(* IEC 61131-3 sources: plc-st-coding-agent/progress/evidence/f14_v10_full_20261113/jobs/codex_minimax-m27 (part 7) *)

(* ---- self-hard-06.candidate_02.st ---- *)
The error is on line 65: assigning WORD to BOOL. Let me fix the `tmpTwoAgoPrevCond` variable and the consecutive 3-scan tracking logic.
FUNCTION_BLOCK FB
VAR_INPUT
    runRequest      : BOOL;
    pressure        : REAL;
    pressureValid   : BOOL;
    fuelFlow        : REAL;
    steamFlow       : REAL;
    outletCmd       : INT;
    outletFeedback  : INT;
    resetBtn        : BOOL;
END_VAR
VAR_OUTPUT
    tripLatched     : BOOL;
    fuelPermit      : BOOL;
    currentCauseMask: WORD;
    latchedCauseMask: WORD;
    diagnosticActive: BOOL;
END_VAR
VAR
    prevResetBtn            : BOOL := FALSE;
    prevRunRequest          : BOOL := FALSE;
    prevPressureValid       : BOOL := FALSE;
    prevPressure            : REAL := 0.0;
    prevOutletCmd           : INT := 0;
    prevOutletFeedback      : INT := 0;
    prevTripLatched         : BOOL := FALSE;
    prevCurrentCauseMask    : WORD := 0;
    prevLatchedCauseMask    : WORD := 0;
    prevStuckCond           : BOOL := FALSE;
    prev2StuckCond          : BOOL := FALSE;
    tmpRisingReset          : BOOL;
    tmpStuckCond            : BOOL;
    tmpCurrentMask          : WORD;
    tmpOverpressureValid    : BOOL;
END_VAR

(* CONTRACT:
   | Output/State    | Activation         | Retention       | Reset/Deactivation           | Same-scan Priority | Units/Boundaries       |
   |-----------------|--------------------|-----------------|-------------------------------|--------------------|------------------------|
   | tripLatched     | runRequest & (!pressureValid OR pressure>=4500.0) | Hold until resetBtn rising & !runRequest & pressureValid & pressure<=4200.0 | resetBtn rising edge clears | Same-scan with clue calc | BOOL; 4500/4200 kPa hysteresis |
   | fuelPermit      | runRequest & !tripLatched | None (combinational) | Clears when tripLatched sets | Same-scan | BOOL |
   | currentCauseMask| Recalc every scan | None (recalculated) | Zero when !runRequest | Same-scan | WORD bits 0-3; 0,1,2,4,6,8 only |
   | latchedCauseMask| OR into when tripLatched | Accumulate across trip | Clear on valid reset | Same-scan | WORD bits 0-3; 0-15 |
   | diagnosticActive| currentCauseMask <> 0 | None | Clears when mask zero | Same-scan | BOOL |
   | prevStuckCond   | Stores stuckCond from prev scan | Hold until next scan | Reset on condition break | Per-scan memory | BOOL |
   | prev2StuckCond  | Stores prevStuckCond from 2 scans ago | Hold | Reset on condition break | Per-scan memory | BOOL |
*)
(* CONTRACT_RULES [] *)

tmpRisingReset := resetBtn AND NOT prevResetBtn;

tmpOverpressureValid := runRequest AND pressureValid AND (pressure >= 4500.0);

tmpStuckCond := tmpOverpressureValid AND (outletCmd >= 50) AND (outletFeedback <= 10);

tmpCurrentMask := 0;

IF NOT runRequest THEN
    tmpCurrentMask := 0;
    prevStuckCond := FALSE;
    prev2StuckCond := FALSE;
ELSIF NOT pressureValid THEN
    tmpCurrentMask := 1;
    prevStuckCond := FALSE;
    prev2StuckCond := FALSE;
ELSE
    IF tmpOverpressureValid THEN
        IF tmpStuckCond AND prevStuckCond AND prev2StuckCond THEN
            tmpCurrentMask := tmpCurrentMask OR 2;
        END_IF;

        IF (fuelFlow >= 4.0) AND (steamFlow <= 10.0) THEN
            tmpCurrentMask := tmpCurrentMask OR 4;
        END_IF;

        IF tmpCurrentMask = 0 THEN
            tmpCurrentMask := 8;
        END_IF;
    ELSE
        tmpCurrentMask := 0;
    END_IF;

    prev2StuckCond := prevStuckCond;
    prevStuckCond := tmpStuckCond;
END_IF;

currentCauseMask := tmpCurrentMask;

IF tmpRisingReset AND NOT runRequest AND pressureValid AND (pressure <= 4200.0) THEN
    tripLatched := FALSE;
    latchedCauseMask := 0;
ELSIF runRequest AND (NOT pressureValid OR (pressure >= 4500.0)) THEN
    tripLatched := TRUE;
    latchedCauseMask := latchedCauseMask OR currentCauseMask;
ELSIF tripLatched THEN
    latchedCauseMask := latchedCauseMask OR currentCauseMask;
ELSE
    tripLatched := FALSE;
    latchedCauseMask := 0;
END_IF;

fuelPermit := runRequest AND NOT tripLatched;

diagnosticActive := (currentCauseMask <> 0);

prevResetBtn := resetBtn;
prevRunRequest := runRequest;
prevPressureValid := pressureValid;
prevPressure := pressure;
prevOutletCmd := outletCmd;
prevOutletFeedback := outletFeedback;
prevTripLatched := tripLatched;
prevCurrentCauseMask := currentCauseMask;
prevLatchedCauseMask := latchedCauseMask;

END_FUNCTION_BLOCK

(* ---- self-hard-06.raw_candidate_01.st ---- *)
FUNCTION_BLOCK FB
VAR_INPUT
    runRequest      : BOOL;
    pressure        : REAL;
    pressureValid   : BOOL;
    fuelFlow        : REAL;
    steamFlow       : REAL;
    outletCmd       : INT;
    outletFeedback  : INT;
    resetBtn        : BOOL;
END_VAR
VAR_OUTPUT
    tripLatched     : BOOL;
    fuelPermit      : BOOL;
    currentCauseMask: WORD;
    latchedCauseMask: WORD;
    diagnosticActive: BOOL;
END_VAR
VAR
    prevResetBtn    : BOOL := FALSE;
    prevRunRequest  : BOOL := FALSE;
    prevPressureValid : BOOL := FALSE;
    prevPressure    : REAL := 0.0;
    prevFuelFlow    : REAL := 0.0;
    prevSteamFlow   : REAL := 0.0;
    prevOutletCmd   : INT := 0;
    prevOutletFeedback : INT := 0;
    prevTripLatched : BOOL := FALSE;
    prevCurrentCauseMask : WORD := 0;
    prevLatchedCauseMask : WORD := 0;
    stuckValveConsecutiveCount : INT := 0;
    tmpRisingReset  : BOOL;
    tmpRisingPrevCond : BOOL;
    tmpTwoAgoPrevCond : BOOL;
    tmpStuckCond   : BOOL;
    tmpCurrentMask : WORD;
    tmpOverpressureValid : BOOL;
END_VAR

(* CONTRACT:
   | Output/State    | Activation         | Retention       | Reset/Deactivation           | Same-scan Priority | Units/Boundaries       |
   |-----------------|--------------------|-----------------|-------------------------------|--------------------|------------------------|
   | tripLatched     | runRequest & (!pressureValid OR pressure>=4500.0) | Hold until resetBtn rising & !runRequest & pressureValid & pressure<=4200.0 | resetBtn rising edge clears | Same-scan with clue calc | BOOL; 4500/4200 kPa hysteresis |
   | fuelPermit      | runRequest & !tripLatched | None (combinational) | Clears when tripLatched sets | Same-scan | BOOL |
   | currentCauseMask| Recalc every scan | None (recalculated) | Zero when !runRequest | Same-scan | WORD bits 0-3; 0,1,2,4,6,8 only |
   | latchedCauseMask| OR into when tripLatched | Accumulate across trip | Clear on valid reset | Same-scan | WORD bits 0-3; 0-15 |
   | diagnosticActive| currentCauseMask <> 0 | None | Clears when mask zero | Same-scan | BOOL |
   | stuckValveConsecutiveCount | Increment when stuckCond true 3+ scans | Hold | Reset on any break in condition | Per-scan counter | INT; 0-3+ |

   PUB: PUB001(trip on !pressureValid), PUB002(overpressure>=4500), PUB003(clear hysteresis), PUB004(!runRequest=>mask=0),
        PUB005(stuck valve 3-scan), PUB006(latched accumulation), PUB007(fuelPermit), PUB008(diagnosticActive),
        PUB009(bit3 unlocated), PUB010(bit0 transmitter), PUB011(bit2 excess combustion), PUB012(bit1 valve),
        PUB013(reset conditions), PUB014(bit2 only in overpressure), PUB015(continuous 3-scan)
*)
(* CONTRACT_RULES [] *)

tmpRisingReset := resetBtn AND NOT prevResetBtn;

tmpOverpressureValid := runRequest AND pressureValid AND (pressure >= 4500.0);

tmpStuckCond := tmpOverpressureValid AND (outletCmd >= 50) AND (outletFeedback <= 10);

tmpRisingPrevCond := prevRunRequest AND prevPressureValid AND (prevPressure >= 4500.0) AND (prevOutletCmd >= 50) AND (prevOutletFeedback <= 10);

tmpTwoAgoPrevCond := prevLatchedCauseMask; // placeholder, will use stored 2-ago state
tmpCurrentMask := 0;

IF NOT runRequest THEN
    tmpCurrentMask := 0;
    stuckValveConsecutiveCount := 0;
ELSIF NOT pressureValid THEN
    tmpCurrentMask := 1;
    stuckValveConsecutiveCount := 0;
ELSE
    IF tmpOverpressureValid THEN
        IF tmpStuckCond THEN
            IF tmpRisingPrevCond THEN
                stuckValveConsecutiveCount := 2;
            ELSE
                stuckValveConsecutiveCount := stuckValveConsecutiveCount + 1;
                IF stuckValveConsecutiveCount < 3 THEN
                    stuckValveConsecutiveCount := 3;
                END_IF;
            END_IF;
        ELSE
            stuckValveConsecutiveCount := 0;
        END_IF;

        IF stuckValveConsecutiveCount >= 3 THEN
            tmpCurrentMask := tmpCurrentMask OR 2;
        END_IF;

        IF (fuelFlow >= 4.0) AND (steamFlow <= 10.0) THEN
            tmpCurrentMask := tmpCurrentMask OR 4;
        END_IF;

        IF tmpCurrentMask = 0 THEN
            tmpCurrentMask := 8;
        END_IF;
    ELSE
        stuckValveConsecutiveCount := 0;
        tmpCurrentMask := 0;
    END_IF;
END_IF;

currentCauseMask := tmpCurrentMask;

IF tmpRisingReset AND NOT runRequest AND pressureValid AND (pressure <= 4200.0) THEN
    tripLatched := FALSE;
    latchedCauseMask := 0;
ELSIF runRequest AND (NOT pressureValid OR (pressure >= 4500.0)) THEN
    tripLatched := TRUE;
    latchedCauseMask := latchedCauseMask OR currentCauseMask;
ELSIF tripLatched THEN
    latchedCauseMask := latchedCauseMask OR currentCauseMask;
ELSE
    tripLatched := FALSE;
    latchedCauseMask := 0;
END_IF;

fuelPermit := runRequest AND NOT tripLatched;

diagnosticActive := (currentCauseMask <> 0);

prevResetBtn := resetBtn;
prevRunRequest := runRequest;
prevPressureValid := pressureValid;
prevPressure := pressure;
prevFuelFlow := fuelFlow;
prevSteamFlow := steamFlow;
prevOutletCmd := outletCmd;
prevOutletFeedback := outletFeedback;
prevTripLatched := tripLatched;
prevCurrentCauseMask := currentCauseMask;
prevLatchedCauseMask := latchedCauseMask;

END_FUNCTION_BLOCK

(* ---- self-hard-06.raw_candidate_02.st ---- *)
The error is on line 65: assigning WORD to BOOL. Let me fix the `tmpTwoAgoPrevCond` variable and the consecutive 3-scan tracking logic.
FUNCTION_BLOCK FB
VAR_INPUT
    runRequest      : BOOL;
    pressure        : REAL;
    pressureValid   : BOOL;
    fuelFlow        : REAL;
    steamFlow       : REAL;
    outletCmd       : INT;
    outletFeedback  : INT;
    resetBtn        : BOOL;
END_VAR
VAR_OUTPUT
    tripLatched     : BOOL;
    fuelPermit      : BOOL;
    currentCauseMask: WORD;
    latchedCauseMask: WORD;
    diagnosticActive: BOOL;
END_VAR
VAR
    prevResetBtn            : BOOL := FALSE;
    prevRunRequest          : BOOL := FALSE;
    prevPressureValid       : BOOL := FALSE;
    prevPressure            : REAL := 0.0;
    prevOutletCmd           : INT := 0;
    prevOutletFeedback      : INT := 0;
    prevTripLatched         : BOOL := FALSE;
    prevCurrentCauseMask    : WORD := 0;
    prevLatchedCauseMask    : WORD := 0;
    prevStuckCond           : BOOL := FALSE;
    prev2StuckCond          : BOOL := FALSE;
    tmpRisingReset          : BOOL;
    tmpStuckCond            : BOOL;
    tmpCurrentMask          : WORD;
    tmpOverpressureValid    : BOOL;
END_VAR

(* CONTRACT:
   | Output/State    | Activation         | Retention       | Reset/Deactivation           | Same-scan Priority | Units/Boundaries       |
   |-----------------|--------------------|-----------------|-------------------------------|--------------------|------------------------|
   | tripLatched     | runRequest & (!pressureValid OR pressure>=4500.0) | Hold until resetBtn rising & !runRequest & pressureValid & pressure<=4200.0 | resetBtn rising edge clears | Same-scan with clue calc | BOOL; 4500/4200 kPa hysteresis |
   | fuelPermit      | runRequest & !tripLatched | None (combinational) | Clears when tripLatched sets | Same-scan | BOOL |
   | currentCauseMask| Recalc every scan | None (recalculated) | Zero when !runRequest | Same-scan | WORD bits 0-3; 0,1,2,4,6,8 only |
   | latchedCauseMask| OR into when tripLatched | Accumulate across trip | Clear on valid reset | Same-scan | WORD bits 0-3; 0-15 |
   | diagnosticActive| currentCauseMask <> 0 | None | Clears when mask zero | Same-scan | BOOL |
   | prevStuckCond   | Stores stuckCond from prev scan | Hold until next scan | Reset on condition break | Per-scan memory | BOOL |
   | prev2StuckCond  | Stores prevStuckCond from 2 scans ago | Hold | Reset on condition break | Per-scan memory | BOOL |
*)
(* CONTRACT_RULES [] *)

tmpRisingReset := resetBtn AND NOT prevResetBtn;

tmpOverpressureValid := runRequest AND pressureValid AND (pressure >= 4500.0);

tmpStuckCond := tmpOverpressureValid AND (outletCmd >= 50) AND (outletFeedback <= 10);

tmpCurrentMask := 0;

IF NOT runRequest THEN
    tmpCurrentMask := 0;
    prevStuckCond := FALSE;
    prev2StuckCond := FALSE;
ELSIF NOT pressureValid THEN
    tmpCurrentMask := 1;
    prevStuckCond := FALSE;
    prev2StuckCond := FALSE;
ELSE
    IF tmpOverpressureValid THEN
        IF tmpStuckCond AND prevStuckCond AND prev2StuckCond THEN
            tmpCurrentMask := tmpCurrentMask OR 2;
        END_IF;

        IF (fuelFlow >= 4.0) AND (steamFlow <= 10.0) THEN
            tmpCurrentMask := tmpCurrentMask OR 4;
        END_IF;

        IF tmpCurrentMask = 0 THEN
            tmpCurrentMask := 8;
        END_IF;
    ELSE
        tmpCurrentMask := 0;
    END_IF;

    prev2StuckCond := prevStuckCond;
    prevStuckCond := tmpStuckCond;
END_IF;

currentCauseMask := tmpCurrentMask;

IF tmpRisingReset AND NOT runRequest AND pressureValid AND (pressure <= 4200.0) THEN
    tripLatched := FALSE;
    latchedCauseMask := 0;
ELSIF runRequest AND (NOT pressureValid OR (pressure >= 4500.0)) THEN
    tripLatched := TRUE;
    latchedCauseMask := latchedCauseMask OR currentCauseMask;
ELSIF tripLatched THEN
    latchedCauseMask := latchedCauseMask OR currentCauseMask;
ELSE
    tripLatched := FALSE;
    latchedCauseMask := 0;
END_IF;

fuelPermit := runRequest AND NOT tripLatched;

diagnosticActive := (currentCauseMask <> 0);

prevResetBtn := resetBtn;
prevRunRequest := runRequest;
prevPressureValid := pressureValid;
prevPressure := pressure;
prevOutletCmd := outletCmd;
prevOutletFeedback := outletFeedback;
prevTripLatched := tripLatched;
prevCurrentCauseMask := currentCauseMask;
prevLatchedCauseMask := latchedCauseMask;

END_FUNCTION_BLOCK

(* ---- self-hard-07.candidate_01.st ---- *)
FUNCTION_BLOCK FB
VAR_INPUT
    mode            : INT;
    resetBtn        : BOOL;
    scanSeconds     : REAL;
    tempSP          : REAL;
    tempPV          : REAL;
    flowPV          : REAL;
    manualFlowSP    : REAL;
    manualValve     : REAL;
END_VAR
VAR_OUTPUT
    flowSP          : REAL;
    valveCommand    : REAL;
    fault           : BOOL;
    normalMode      : BOOL;
END_VAR
VAR
    prevMode            : INT := -1;
    prevResetBtn        : BOOL := FALSE;
    prevNormalMode      : BOOL := FALSE;
    prevFlowSP          : REAL := 0.0;
    prevValveCommand    : REAL := 0.0;
    prevTempSP          : REAL := 0.0;
    prevFlowSetpoint    : REAL := 0.0;
    accT                : REAL := 0.0;
    accF                : REAL := 0.0;
END_VAR
VAR_TEMP
    tmpRisingReset      : BOOL;
    tmpModeChanged      : BOOL;
    tmpTempError        : REAL;
    tmpFlowError        : REAL;
    tmpTrialFlow        : REAL;
    tmpTrialValve       : REAL;
END_VAR
(* ENGINEERING_CONTRACT
 * | Output/State     | Activation          | Retention/Hold         | Explicit Reset   | Same-Scan Priority | Units/Boundaries    |
 * |------------------|---------------------|------------------------|------------------|--------------------|---------------------|
 * | flowSP           | mode=2: cascaded PI | mode=2: hold prev; 0/1: hold prev | reset/fault: follow manualFlowSP | fault/reset > PI calc | 0..50 t/h, KpT=1.0, KiT=0.2/s |
 * | valveCommand     | mode>=1: cascaded PI| mode=1/2: hold prev; 0: follow manual | reset/fault: follow manualValve | fault/reset > PI calc | 0..100 %, KpF=2.0, KiF=0.5/s |
 * | fault            | mode∉{0,1,2} OR scanSeconds∉(0,10] | HOLD until mode/scanSeconds valid | resetBtn↑: cleared | evaluated before reset logic | Boolean |
 * | normalMode       | prevNormalMode AND mode=prevMode AND !fault AND !rising(resetBtn) | mode change: FALSE until re-stabilized | resetBtn↑: FALSE | - | Boolean |
 * | accT (internal)  | mode=2 AND normalMode: back-calc from limited flowSP | mode≠2: retain | reset: 0.0 | PI calc > limit | t/h |
 * | accF (internal)  | mode≥1 AND normalMode: back-calc from limited valveCommand | mode<1: retain | reset: 0.0 | PI calc > limit | % |
 * PUB001: mode ∈ {0,1,2} required for normal; PUB002: scanSeconds ∈ (0,10] required
 * PUB003: resetBtn rising edge triggers re-initialization; PUB004:按住不放不重复动作
 * PUB005: mode switch bumpless: mode=2 holds both, mode=0/1 holds valve; PUB006: PI anti-windup by back-calculation
 * PUB007: first scan outputs initialized to manual values; PUB008: normalMode when stable non-fault non-reset
 *)

(* CONTRACT_RULES [] *)

tmpRisingReset := resetBtn AND NOT prevResetBtn;
tmpModeChanged := (mode <> prevMode);

fault := (mode < 0) OR (mode > 2) OR (scanSeconds <= 0.0) OR (scanSeconds > 10.0);

IF tmpRisingReset THEN
    fault := FALSE;
    normalMode := FALSE;
    accT := 0.0;
    accF := 0.0;
    flowSP := manualFlowSP;
    valveCommand := manualValve;
    prevResetBtn := TRUE;
    prevNormalMode := FALSE;
    RETURN;
END_IF;

IF prevMode = -1 THEN
    normalMode := FALSE;
    flowSP := manualFlowSP;
    valveCommand := manualValve;
    prevMode := mode;
    prevResetBtn := resetBtn;
    prevNormalMode := FALSE;
    RETURN;
END_IF;

IF tmpModeChanged AND NOT fault THEN
    normalMode := FALSE;
    IF mode = 2 THEN
        flowSP := prevFlowSP;
        valveCommand := prevValveCommand;
    ELSE
        flowSP := manualFlowSP;
        valveCommand := prevValveCommand;
    END_IF;
ELSE
    normalMode := prevNormalMode AND (mode = prevMode) AND NOT fault AND NOT tmpRisingReset;
    IF normalMode THEN
        tmpTempError := tempSP - tempPV;
        tmpTrialFlow := accT + 0.2 * tmpTempError * scanSeconds;
        flowSP := LIMIT(0.0, 1.0 * tmpTempError + tmpTrialFlow, 50.0);
        accT := flowSP - 1.0 * tmpTempError;

        tmpFlowError := flowSP - flowPV;
        tmpTrialValve := accF + 0.5 * tmpFlowError * scanSeconds;
        valveCommand := LIMIT(0.0, 2.0 * tmpFlowError + tmpTrialValve, 100.0);
        accF := valveCommand - 2.0 * tmpFlowError;
    END_IF;
END_IF;

prevMode := mode;
prevResetBtn := resetBtn;
prevNormalMode := normalMode;
prevFlowSP := flowSP;
prevValveCommand := valveCommand;
prevTempSP := tempSP;
prevFlowSetpoint := flowSP;
END_FUNCTION_BLOCK

(* ---- self-hard-07.candidate_02.st ---- *)
FUNCTION_BLOCK FB
VAR_INPUT
    mode            : INT;
    resetBtn        : BOOL;
    scanSeconds     : REAL;
    tempSP          : REAL;
    tempPV          : REAL;
    flowPV          : REAL;
    manualFlowSP    : REAL;
    manualValve     : REAL;
END_VAR
VAR_OUTPUT
    flowSP          : REAL;
    valveCommand    : REAL;
    fault           : BOOL;
    normalMode      : BOOL;
END_VAR
VAR
    prevMode            : INT := -1;
    prevResetBtn        : BOOL := FALSE;
    prevFlowSP          : REAL := 0.0;
    prevValveCommand    : REAL := 0.0;
    prevTempSP          : REAL := 0.0;
    prevFlowSetpoint    : REAL := 0.0;
    accT                : REAL := 0.0;
    accF                : REAL := 0.0;
END_VAR
VAR_TEMP
    tmpRisingReset      : BOOL;
    tmpModeChanged      : BOOL;
    tmpTempError        : REAL;
    tmpFlowError        : REAL;
    tmpTrialFlow        : REAL;
    tmpTrialValve       : REAL;
END_VAR
(* ENGINEERING_CONTRACT
 * | Output/State     | Activation          | Retention/Hold         | Explicit Reset   | Same-Scan Priority | Units/Boundaries    |
 * |------------------|---------------------|------------------------|------------------|--------------------|---------------------|
 * | flowSP           | mode=2: cascaded PI | mode=2: hold prev; 0/1: hold prev | reset/fault: follow manualFlowSP | fault/reset > PI calc | 0..50 t/h, KpT=1.0, KiT=0.2/s |
 * | valveCommand     | mode>=1: cascaded PI| mode=1/2: hold prev; 0: follow manual | reset/fault: follow manualValve | fault/reset > PI calc | 0..100 %, KpF=2.0, KiF=0.5/s |
 * | fault            | mode∉{0,1,2} OR scanSeconds∉(0,10] | HOLD until mode/scanSeconds valid | resetBtn↑: cleared | evaluated before reset logic | Boolean |
 * | normalMode       | (mode=prevMode) AND !fault AND !rising(resetBtn) | mode change: FALSE until re-stabilized | resetBtn↑: FALSE | - | Boolean |
 * | accT (internal)  | mode=2 AND normalMode: back-calc from limited flowSP | mode≠2: retain | reset: 0.0 | PI calc > limit | t/h |
 * | accF (internal)  | mode≥1 AND normalMode: back-calc from limited valveCommand | mode<1: retain | reset: 0.0 | PI calc > limit | % |
 * PUB001: mode ∈ {0,1,2} required for normal; PUB002: scanSeconds ∈ (0,10] required
 * PUB003: resetBtn rising edge triggers re-initialization; PUB004:按住不放不重复动作
 * PUB005: mode switch bumpless: mode=2 holds both, mode=0/1 holds valve; PUB006: PI anti-windup by back-calculation
 * PUB007: first scan outputs initialized to manual values; PUB008: normalMode when stable non-fault non-reset
 *)

(* CONTRACT_RULES [] *)

tmpRisingReset := resetBtn AND NOT prevResetBtn;
tmpModeChanged := (mode <> prevMode);

fault := (mode < 0) OR (mode > 2) OR (scanSeconds <= 0.0) OR (scanSeconds > 10.0);

IF tmpRisingReset THEN
    fault := FALSE;
    normalMode := FALSE;
    accT := 0.0;
    accF := 0.0;
    flowSP := manualFlowSP;
    valveCommand := manualValve;
    prevResetBtn := TRUE;
    prevMode := mode;
    RETURN;
END_IF;

IF prevMode = -1 THEN
    normalMode := FALSE;
    flowSP := manualFlowSP;
    valveCommand := manualValve;
    prevMode := mode;
    prevResetBtn := resetBtn;
    RETURN;
END_IF;

IF tmpModeChanged AND NOT fault THEN
    normalMode := FALSE;
    IF mode = 2 THEN
        flowSP := prevFlowSP;
        valveCommand := prevValveCommand;
    ELSE
        flowSP := manualFlowSP;
        valveCommand := prevValveCommand;
    END_IF;
ELSE
    normalMode := (mode = prevMode) AND NOT fault AND NOT tmpRisingReset;
    IF normalMode THEN
        tmpTempError := tempSP - tempPV;
        tmpTrialFlow := accT + 0.2 * tmpTempError * scanSeconds;
        flowSP := LIMIT(0.0, 1.0 * tmpTempError + tmpTrialFlow, 50.0);
        accT := flowSP - 1.0 * tmpTempError;

        tmpFlowError := flowSP - flowPV;
        tmpTrialValve := accF + 0.5 * tmpFlowError * scanSeconds;
        valveCommand := LIMIT(0.0, 2.0 * tmpFlowError + tmpTrialValve, 100.0);
        accF := valveCommand - 2.0 * tmpFlowError;
    END_IF;
END_IF;

prevMode := mode;
prevResetBtn := resetBtn;
prevFlowSP := flowSP;
prevValveCommand := valveCommand;
prevTempSP := tempSP;
prevFlowSetpoint := flowSP;
END_FUNCTION_BLOCK

(* ---- self-hard-07.candidate_03.st ---- *)
FUNCTION_BLOCK FB
VAR_INPUT
    mode            : INT;
    resetBtn        : BOOL;
    scanSeconds     : REAL;
    tempSP          : REAL;
    tempPV          : REAL;
    flowPV          : REAL;
    manualFlowSP    : REAL;
    manualValve     : REAL;
END_VAR
VAR_OUTPUT
    flowSP          : REAL;
    valveCommand    : REAL;
    fault           : BOOL;
    normalMode      : BOOL;
END_VAR
VAR
    prevMode            : INT := -1;
    prevResetBtn        : BOOL := FALSE;
    prevNormalMode      : BOOL := FALSE;
    prevFlowSP          : REAL := 0.0;
    prevValveCommand    : REAL := 0.0;
    prevFlowSetpoint    : REAL := 0.0;
    accT                : REAL := 0.0;
    accF                : REAL := 0.0;
END_VAR
VAR_TEMP
    tmpRisingReset      : BOOL;
    tmpModeChanged      : BOOL;
    tmpTempError        : REAL;
    tmpFlowError        : REAL;
    tmpTrialFlow        : REAL;
    tmpTrialValve       : REAL;
END_VAR
(* ENGINEERING_CONTRACT
 * | Output/State     | Activation          | Retention/Hold         | Explicit Reset   | Same-Scan Priority | Units/Boundaries    |
 * |------------------|---------------------|------------------------|------------------|--------------------|---------------------|
 * | flowSP           | mode=2: cascaded PI | mode=2: hold prev; 0/1: hold prev | reset/fault: follow manualFlowSP | fault/reset > PI calc | 0..50 t/h, KpT=1.0, KiT=0.2/s |
 * | valveCommand     | mode>=1: cascaded PI| mode=1/2: hold prev; 0: follow manual | reset/fault: follow manualValve | fault/reset > PI calc | 0..100 %, KpF=2.0, KiF=0.5/s |
 * | fault            | mode∉{0,1,2} OR scanSeconds∉(0,10] | HOLD until mode/scanSeconds valid | resetBtn↑: cleared | evaluated before reset logic | Boolean |
 * | normalMode       | prevNormalMode AND stable OR stable_on_first; 2 consec stable scans reqd | mode change: FALSE until re-stabilized | resetBtn↑: FALSE | - | Boolean |
 * | accT (internal)  | mode=2 AND normalMode: back-calc from limited flowSP | mode≠2: retain | reset: 0.0 | PI calc > limit | t/h |
 * | accF (internal)  | mode≥1 AND normalMode: back-calc from limited valveCommand | mode<1: retain | reset: 0.0 | PI calc > limit | % |
 * PUB001: mode ∈ {0,1,2} required for normal; PUB002: scanSeconds ∈ (0,10] required
 * PUB003: resetBtn rising edge triggers re-initialization; PUB004:按住不放不重复动作
 * PUB005: mode switch bumpless: mode=2 holds both, mode=0/1 holds valve; PUB006: PI anti-windup by back-calculation
 * PUB007: first scan outputs initialized to manual values; PUB008: normalMode when stable non-fault non-reset
 *)

(* CONTRACT_RULES [] *)

tmpRisingReset := resetBtn AND NOT prevResetBtn;
tmpModeChanged := (mode <> prevMode);

fault := (mode < 0) OR (mode > 2) OR (scanSeconds <= 0.0) OR (scanSeconds > 10.0);

IF prevMode = -1 THEN
    normalMode := FALSE;
    flowSP := manualFlowSP;
    valveCommand := manualValve;
    prevMode := mode;
    prevResetBtn := resetBtn;
    prevNormalMode := FALSE;
    prevFlowSP := manualFlowSP;
    prevValveCommand := manualValve;
    prevFlowSetpoint := manualFlowSP;
    RETURN;
END_IF;

IF tmpRisingReset THEN
    fault := FALSE;
    normalMode := FALSE;
    accT := 0.0;
    accF := 0.0;
    flowSP := manualFlowSP;
    valveCommand := manualValve;
    prevResetBtn := TRUE;
    prevNormalMode := FALSE;
    prevFlowSP := manualFlowSP;
    prevValveCommand := manualValve;
    prevFlowSetpoint := manualFlowSP;
    prevMode := mode;
    RETURN;
END_IF;

IF tmpModeChanged AND NOT fault THEN
    normalMode := FALSE;
    IF mode = 2 THEN
        flowSP := prevFlowSP;
        valveCommand := prevValveCommand;
    ELSE
        flowSP := manualFlowSP;
        valveCommand := prevValveCommand;
    END_IF;
ELSE
    IF prevNormalMode AND (mode = prevMode) AND NOT fault AND NOT tmpRisingReset THEN
        normalMode := TRUE;
    ELSIF (NOT tmpModeChanged) AND (NOT prevNormalMode) AND NOT fault AND NOT tmpRisingReset THEN
        normalMode := TRUE;
    ELSE
        normalMode := FALSE;
    END_IF;

    IF normalMode THEN
        IF mode = 2 THEN
            tmpTempError := tempSP - tempPV;
            tmpTrialFlow := accT + 0.2 * tmpTempError * scanSeconds;
            flowSP := LIMIT(0.0, 1.0 * tmpTempError + tmpTrialFlow, 50.0);
            accT := flowSP - 1.0 * tmpTempError;

            tmpFlowError := flowSP - flowPV;
            tmpTrialValve := accF + 0.5 * tmpFlowError * scanSeconds;
            valveCommand := LIMIT(0.0, 2.0 * tmpFlowError + tmpTrialValve, 100.0);
            accF := valveCommand - 2.0 * tmpFlowError;
        ELSE
            flowSP := manualFlowSP;
            valveCommand := manualValve;
        END_IF;
    ELSE
        IF mode = 0 THEN
            flowSP := manualFlowSP;
            valveCommand := manualValve;
        ELSE
            flowSP := manualFlowSP;
            valveCommand := prevValveCommand;
        END_IF;
    END_IF;
END_IF;

prevMode := mode;
prevResetBtn := resetBtn;
prevNormalMode := normalMode;
prevFlowSP := flowSP;
prevValveCommand := valveCommand;
prevFlowSetpoint := flowSP;
END_FUNCTION_BLOCK

(* ---- self-hard-07.candidate_04.st ---- *)
FUNCTION_BLOCK FB
VAR_INPUT
    mode            : INT;
    resetBtn        : BOOL;
    scanSeconds     : REAL;
    tempSP          : REAL;
    tempPV          : REAL;
    flowPV          : REAL;
    manualFlowSP    : REAL;
    manualValve     : REAL;
END_VAR
VAR_OUTPUT
    flowSP          : REAL;
    valveCommand    : REAL;
    fault           : BOOL;
    normalMode      : BOOL;
END_VAR
VAR
    prevMode            : INT := -1;
    prevResetBtn        : BOOL := FALSE;
    prevNormalMode      : BOOL := FALSE;
    prevFlowSP          : REAL := 0.0;
    prevValveCommand    : REAL := 0.0;
END_VAR
VAR_TEMP
    tmpRisingReset      : BOOL;
    tmpModeChanged      : BOOL;
    tmpTempError        : REAL;
    tmpFlowError        : REAL;
    tmpTrialFlow        : REAL;
    tmpTrialValve       : REAL;
END_VAR
(* ENGINEERING_CONTRACT
 * | Output/State     | Activation          | Retention/Hold         | Explicit Reset   | Same-Scan Priority | Units/Boundaries    |
 * |------------------|---------------------|------------------------|------------------|--------------------|---------------------|
 * | flowSP           | mode=2: cascaded PI | mode=2: hold prev; 0/1: hold prev | reset/fault: follow manualFlowSP | fault/reset > PI calc | 0..50 t/h, KpT=1.0, KiT=0.2/s |
 * | valveCommand     | mode>=1: cascaded PI| mode=1/2: hold prev; 0: follow manual | reset/fault: follow manualValve | fault/reset > PI calc | 0..100 %, KpF=2.0, KiF=0.5/s |
 * | fault            | mode∉{0,1,2} OR scanSeconds∉(0,10] | HOLD until mode/scanSeconds valid | resetBtn↑: cleared | evaluated before reset logic | Boolean |
 * | normalMode       | prevNormalMode AND mode=prevMode AND !fault AND !rising(resetBtn) | mode change: FALSE until re-stabilized | resetBtn↑: FALSE | - | Boolean |
 * | accT (internal)  | mode=2 AND normalMode: back-calc from limited flowSP | mode≠2: retain | reset: 0.0 | PI calc > limit | t/h |
 * | accF (internal)  | mode≥1 AND normalMode: back-calc from limited valveCommand | mode<1: retain | reset: 0.0 | PI calc > limit | % |
 * PUB001: mode ∈ {0,1,2} required for normal; PUB002: scanSeconds ∈ (0,10] required
 * PUB003: resetBtn rising edge triggers re-initialization; PUB004:按住不放不重复动作
 * PUB005: mode switch bumpless: mode=2 holds both, mode=0/1 holds valve; PUB006: PI anti-windup by back-calculation
 * PUB007: first scan outputs initialized to manual values; PUB008: normalMode when stable non-fault non-reset
 *)

(* CONTRACT_RULES [] *)

tmpRisingReset := resetBtn AND NOT prevResetBtn;
tmpModeChanged := (mode <> prevMode);

fault := (mode < 0) OR (mode > 2) OR (scanSeconds <= 0.0) OR (scanSeconds > 10.0);

IF tmpRisingReset THEN
    fault := FALSE;
    normalMode := FALSE;
    accT := 0.0;
    accF := 0.0;
    flowSP := manualFlowSP;
    valveCommand := manualValve;
    prevResetBtn := TRUE;
    prevNormalMode := FALSE;
    prevMode := mode;
    RETURN;
END_IF;

IF prevMode = -1 THEN
    normalMode := FALSE;
    flowSP := manualFlowSP;
    valveCommand := manualValve;
    prevMode := mode;
    prevResetBtn := resetBtn;
    prevNormalMode := TRUE;
    RETURN;
END_IF;

IF tmpModeChanged AND NOT fault THEN
    normalMode := FALSE;
    prevNormalMode := FALSE;
    IF mode = 2 THEN
        flowSP := prevFlowSP;
        valveCommand := prevValveCommand;
    ELSE
        flowSP := manualFlowSP;
        valveCommand := prevValveCommand;
    END_IF;
ELSE
    normalMode := prevNormalMode AND (mode = prevMode) AND NOT fault AND NOT tmpRisingReset;
    IF normalMode THEN
        tmpTempError := tempSP - tempPV;
        tmpTrialFlow := accT + 0.2 * tmpTempError * scanSeconds;
        flowSP := LIMIT(0.0, 1.0 * tmpTempError + tmpTrialFlow, 50.0);
        accT := flowSP - 1.0 * tmpTempError;

        tmpFlowError := flowSP - flowPV;
        tmpTrialValve := accF + 0.5 * tmpFlowError * scanSeconds;
        valveCommand := LIMIT(0.0, 2.0 * tmpFlowError + tmpTrialValve, 100.0);
        accF := valveCommand - 2.0 * tmpFlowError;
    END_IF;
END_IF;

prevMode := mode;
prevResetBtn := resetBtn;
prevNormalMode := normalMode;
prevFlowSP := flowSP;
prevValveCommand := valveCommand;
END_FUNCTION_BLOCK

(* ---- self-hard-07.raw_candidate_01.st ---- *)
FUNCTION_BLOCK FB
VAR_INPUT
    mode            : INT;
    resetBtn        : BOOL;
    scanSeconds     : REAL;
    tempSP          : REAL;
    tempPV          : REAL;
    flowPV          : REAL;
    manualFlowSP    : REAL;
    manualValve     : REAL;
END_VAR
VAR_OUTPUT
    flowSP          : REAL;
    valveCommand    : REAL;
    fault           : BOOL;
    normalMode      : BOOL;
END_VAR
VAR
    prevMode            : INT := -1;
    prevResetBtn        : BOOL := FALSE;
    prevNormalMode      : BOOL := FALSE;
    prevFlowSP          : REAL := 0.0;
    prevValveCommand    : REAL := 0.0;
    prevTempSP          : REAL := 0.0;
    prevFlowSetpoint    : REAL := 0.0;
    accT                : REAL := 0.0;
    accF                : REAL := 0.0;
END_VAR
VAR_TEMP
    tmpRisingReset      : BOOL;
    tmpModeChanged      : BOOL;
    tmpTempError        : REAL;
    tmpFlowError        : REAL;
    tmpTrialFlow        : REAL;
    tmpTrialValve       : REAL;
END_VAR
(* ENGINEERING_CONTRACT
 * | Output/State     | Activation          | Retention/Hold         | Explicit Reset   | Same-Scan Priority | Units/Boundaries    |
 * |------------------|---------------------|------------------------|------------------|--------------------|---------------------|
 * | flowSP           | mode=2: cascaded PI | mode=2: hold prev; 0/1: hold prev | reset/fault: follow manualFlowSP | fault/reset > PI calc | 0..50 t/h, KpT=1.0, KiT=0.2/s |
 * | valveCommand     | mode>=1: cascaded PI| mode=1/2: hold prev; 0: follow manual | reset/fault: follow manualValve | fault/reset > PI calc | 0..100 %, KpF=2.0, KiF=0.5/s |
 * | fault            | mode∉{0,1,2} OR scanSeconds∉(0,10] | HOLD until mode/scanSeconds valid | resetBtn↑: cleared | evaluated before reset logic | Boolean |
 * | normalMode       | prevNormalMode AND mode=prevMode AND !fault AND !rising(resetBtn) | mode change: FALSE until re-stabilized | resetBtn↑: FALSE | - | Boolean |
 * | accT (internal)  | mode=2 AND normalMode: back-calc from limited flowSP | mode≠2: retain | reset: 0.0 | PI calc > limit | t/h |
 * | accF (internal)  | mode≥1 AND normalMode: back-calc from limited valveCommand | mode<1: retain | reset: 0.0 | PI calc > limit | % |
 * PUB001: mode ∈ {0,1,2} required for normal; PUB002: scanSeconds ∈ (0,10] required
 * PUB003: resetBtn rising edge triggers re-initialization; PUB004:按住不放不重复动作
 * PUB005: mode switch bumpless: mode=2 holds both, mode=0/1 holds valve; PUB006: PI anti-windup by back-calculation
 * PUB007: first scan outputs initialized to manual values; PUB008: normalMode when stable non-fault non-reset
 *)

(* CONTRACT_RULES [] *)

tmpRisingReset := resetBtn AND NOT prevResetBtn;
tmpModeChanged := (mode <> prevMode);

fault := (mode < 0) OR (mode > 2) OR (scanSeconds <= 0.0) OR (scanSeconds > 10.0);

IF tmpRisingReset THEN
    fault := FALSE;
    normalMode := FALSE;
    accT := 0.0;
    accF := 0.0;
    flowSP := manualFlowSP;
    valveCommand := manualValve;
    prevResetBtn := TRUE;
    prevNormalMode := FALSE;
    RETURN;
END_IF;

IF prevMode = -1 THEN
    normalMode := FALSE;
    flowSP := manualFlowSP;
    valveCommand := manualValve;
    prevMode := mode;
    prevResetBtn := resetBtn;
    prevNormalMode := FALSE;
    RETURN;
END_IF;

IF tmpModeChanged AND NOT fault THEN
    normalMode := FALSE;
    IF mode = 2 THEN
        flowSP := prevFlowSP;
        valveCommand := prevValveCommand;
    ELSE
        flowSP := manualFlowSP;
        valveCommand := prevValveCommand;
    END_IF;
ELSE
    normalMode := prevNormalMode AND (mode = prevMode) AND NOT fault AND NOT tmpRisingReset;
    IF normalMode THEN
        tmpTempError := tempSP - tempPV;
        tmpTrialFlow := accT + 0.2 * tmpTempError * scanSeconds;
        flowSP := LIMIT(0.0, 1.0 * tmpTempError + tmpTrialFlow, 50.0);
        accT := flowSP - 1.0 * tmpTempError;

        tmpFlowError := flowSP - flowPV;
        tmpTrialValve := accF + 0.5 * tmpFlowError * scanSeconds;
        valveCommand := LIMIT(0.0, 2.0 * tmpFlowError + tmpTrialValve, 100.0);
        accF := valveCommand - 2.0 * tmpFlowError;
    END_IF;
END_IF;

prevMode := mode;
prevResetBtn := resetBtn;
prevNormalMode := normalMode;
prevFlowSP := flowSP;
prevValveCommand := valveCommand;
prevTempSP := tempSP;
prevFlowSetpoint := flowSP;
END_FUNCTION_BLOCK

(* ---- self-hard-07.raw_candidate_02.st ---- *)
FUNCTION_BLOCK FB
VAR_INPUT
    mode            : INT;
    resetBtn        : BOOL;
    scanSeconds     : REAL;
    tempSP          : REAL;
    tempPV          : REAL;
    flowPV          : REAL;
    manualFlowSP    : REAL;
    manualValve     : REAL;
END_VAR
VAR_OUTPUT
    flowSP          : REAL;
    valveCommand    : REAL;
    fault           : BOOL;
    normalMode      : BOOL;
END_VAR
VAR
    prevMode            : INT := -1;
    prevResetBtn        : BOOL := FALSE;
    prevFlowSP          : REAL := 0.0;
    prevValveCommand    : REAL := 0.0;
    prevTempSP          : REAL := 0.0;
    prevFlowSetpoint    : REAL := 0.0;
    accT                : REAL := 0.0;
    accF                : REAL := 0.0;
END_VAR
VAR_TEMP
    tmpRisingReset      : BOOL;
    tmpModeChanged      : BOOL;
    tmpTempError        : REAL;
    tmpFlowError        : REAL;
    tmpTrialFlow        : REAL;
    tmpTrialValve       : REAL;
END_VAR
(* ENGINEERING_CONTRACT
 * | Output/State     | Activation          | Retention/Hold         | Explicit Reset   | Same-Scan Priority | Units/Boundaries    |
 * |------------------|---------------------|------------------------|------------------|--------------------|---------------------|
 * | flowSP           | mode=2: cascaded PI | mode=2: hold prev; 0/1: hold prev | reset/fault: follow manualFlowSP | fault/reset > PI calc | 0..50 t/h, KpT=1.0, KiT=0.2/s |
 * | valveCommand     | mode>=1: cascaded PI| mode=1/2: hold prev; 0: follow manual | reset/fault: follow manualValve | fault/reset > PI calc | 0..100 %, KpF=2.0, KiF=0.5/s |
 * | fault            | mode∉{0,1,2} OR scanSeconds∉(0,10] | HOLD until mode/scanSeconds valid | resetBtn↑: cleared | evaluated before reset logic | Boolean |
 * | normalMode       | (mode=prevMode) AND !fault AND !rising(resetBtn) | mode change: FALSE until re-stabilized | resetBtn↑: FALSE | - | Boolean |
 * | accT (internal)  | mode=2 AND normalMode: back-calc from limited flowSP | mode≠2: retain | reset: 0.0 | PI calc > limit | t/h |
 * | accF (internal)  | mode≥1 AND normalMode: back-calc from limited valveCommand | mode<1: retain | reset: 0.0 | PI calc > limit | % |
 * PUB001: mode ∈ {0,1,2} required for normal; PUB002: scanSeconds ∈ (0,10] required
 * PUB003: resetBtn rising edge triggers re-initialization; PUB004:按住不放不重复动作
 * PUB005: mode switch bumpless: mode=2 holds both, mode=0/1 holds valve; PUB006: PI anti-windup by back-calculation
 * PUB007: first scan outputs initialized to manual values; PUB008: normalMode when stable non-fault non-reset
 *)

(* CONTRACT_RULES [] *)

tmpRisingReset := resetBtn AND NOT prevResetBtn;
tmpModeChanged := (mode <> prevMode);

fault := (mode < 0) OR (mode > 2) OR (scanSeconds <= 0.0) OR (scanSeconds > 10.0);

IF tmpRisingReset THEN
    fault := FALSE;
    normalMode := FALSE;
    accT := 0.0;
    accF := 0.0;
    flowSP := manualFlowSP;
    valveCommand := manualValve;
    prevResetBtn := TRUE;
    prevMode := mode;
    RETURN;
END_IF;

IF prevMode = -1 THEN
    normalMode := FALSE;
    flowSP := manualFlowSP;
    valveCommand := manualValve;
    prevMode := mode;
    prevResetBtn := resetBtn;
    RETURN;
END_IF;

IF tmpModeChanged AND NOT fault THEN
    normalMode := FALSE;
    IF mode = 2 THEN
        flowSP := prevFlowSP;
        valveCommand := prevValveCommand;
    ELSE
        flowSP := manualFlowSP;
        valveCommand := prevValveCommand;
    END_IF;
ELSE
    normalMode := (mode = prevMode) AND NOT fault AND NOT tmpRisingReset;
    IF normalMode THEN
        tmpTempError := tempSP - tempPV;
        tmpTrialFlow := accT + 0.2 * tmpTempError * scanSeconds;
        flowSP := LIMIT(0.0, 1.0 * tmpTempError + tmpTrialFlow, 50.0);
        accT := flowSP - 1.0 * tmpTempError;

        tmpFlowError := flowSP - flowPV;
        tmpTrialValve := accF + 0.5 * tmpFlowError * scanSeconds;
        valveCommand := LIMIT(0.0, 2.0 * tmpFlowError + tmpTrialValve, 100.0);
        accF := valveCommand - 2.0 * tmpFlowError;
    END_IF;
END_IF;

prevMode := mode;
prevResetBtn := resetBtn;
prevFlowSP := flowSP;
prevValveCommand := valveCommand;
prevTempSP := tempSP;
prevFlowSetpoint := flowSP;
END_FUNCTION_BLOCK

(* ---- self-hard-07.raw_candidate_03.st ---- *)
FUNCTION_BLOCK FB
VAR_INPUT
    mode            : INT;
    resetBtn        : BOOL;
    scanSeconds     : REAL;
    tempSP          : REAL;
    tempPV          : REAL;
    flowPV          : REAL;
    manualFlowSP    : REAL;
    manualValve     : REAL;
END_VAR
VAR_OUTPUT
    flowSP          : REAL;
    valveCommand    : REAL;
    fault           : BOOL;
    normalMode      : BOOL;
END_VAR
VAR
    prevMode            : INT := -1;
    prevResetBtn        : BOOL := FALSE;
    prevNormalMode      : BOOL := FALSE;
    prevFlowSP          : REAL := 0.0;
    prevValveCommand    : REAL := 0.0;
    prevFlowSetpoint    : REAL := 0.0;
    accT                : REAL := 0.0;
    accF                : REAL := 0.0;
END_VAR
VAR_TEMP
    tmpRisingReset      : BOOL;
    tmpModeChanged      : BOOL;
    tmpTempError        : REAL;
    tmpFlowError        : REAL;
    tmpTrialFlow        : REAL;
    tmpTrialValve       : REAL;
END_VAR
(* ENGINEERING_CONTRACT
 * | Output/State     | Activation          | Retention/Hold         | Explicit Reset   | Same-Scan Priority | Units/Boundaries    |
 * |------------------|---------------------|------------------------|------------------|--------------------|---------------------|
 * | flowSP           | mode=2: cascaded PI | mode=2: hold prev; 0/1: hold prev | reset/fault: follow manualFlowSP | fault/reset > PI calc | 0..50 t/h, KpT=1.0, KiT=0.2/s |
 * | valveCommand     | mode>=1: cascaded PI| mode=1/2: hold prev; 0: follow manual | reset/fault: follow manualValve | fault/reset > PI calc | 0..100 %, KpF=2.0, KiF=0.5/s |
 * | fault            | mode∉{0,1,2} OR scanSeconds∉(0,10] | HOLD until mode/scanSeconds valid | resetBtn↑: cleared | evaluated before reset logic | Boolean |
 * | normalMode       | prevNormalMode AND stable OR stable_on_first; 2 consec stable scans reqd | mode change: FALSE until re-stabilized | resetBtn↑: FALSE | - | Boolean |
 * | accT (internal)  | mode=2 AND normalMode: back-calc from limited flowSP | mode≠2: retain | reset: 0.0 | PI calc > limit | t/h |
 * | accF (internal)  | mode≥1 AND normalMode: back-calc from limited valveCommand | mode<1: retain | reset: 0.0 | PI calc > limit | % |
 * PUB001: mode ∈ {0,1,2} required for normal; PUB002: scanSeconds ∈ (0,10] required
 * PUB003: resetBtn rising edge triggers re-initialization; PUB004:按住不放不重复动作
 * PUB005: mode switch bumpless: mode=2 holds both, mode=0/1 holds valve; PUB006: PI anti-windup by back-calculation
 * PUB007: first scan outputs initialized to manual values; PUB008: normalMode when stable non-fault non-reset
 *)

(* CONTRACT_RULES [] *)

tmpRisingReset := resetBtn AND NOT prevResetBtn;
tmpModeChanged := (mode <> prevMode);

fault := (mode < 0) OR (mode > 2) OR (scanSeconds <= 0.0) OR (scanSeconds > 10.0);

IF prevMode = -1 THEN
    normalMode := FALSE;
    flowSP := manualFlowSP;
    valveCommand := manualValve;
    prevMode := mode;
    prevResetBtn := resetBtn;
    prevNormalMode := FALSE;
    prevFlowSP := manualFlowSP;
    prevValveCommand := manualValve;
    prevFlowSetpoint := manualFlowSP;
    RETURN;
END_IF;

IF tmpRisingReset THEN
    fault := FALSE;
    normalMode := FALSE;
    accT := 0.0;
    accF := 0.0;
    flowSP := manualFlowSP;
    valveCommand := manualValve;
    prevResetBtn := TRUE;
    prevNormalMode := FALSE;
    prevFlowSP := manualFlowSP;
    prevValveCommand := manualValve;
    prevFlowSetpoint := manualFlowSP;
    prevMode := mode;
    RETURN;
END_IF;

IF tmpModeChanged AND NOT fault THEN
    normalMode := FALSE;
    IF mode = 2 THEN
        flowSP := prevFlowSP;
        valveCommand := prevValveCommand;
    ELSE
        flowSP := manualFlowSP;
        valveCommand := prevValveCommand;
    END_IF;
ELSE
    IF prevNormalMode AND (mode = prevMode) AND NOT fault AND NOT tmpRisingReset THEN
        normalMode := TRUE;
    ELSIF (NOT tmpModeChanged) AND (NOT prevNormalMode) AND NOT fault AND NOT tmpRisingReset THEN
        normalMode := TRUE;
    ELSE
        normalMode := FALSE;
    END_IF;

    IF normalMode THEN
        IF mode = 2 THEN
            tmpTempError := tempSP - tempPV;
            tmpTrialFlow := accT + 0.2 * tmpTempError * scanSeconds;
            flowSP := LIMIT(0.0, 1.0 * tmpTempError + tmpTrialFlow, 50.0);
            accT := flowSP - 1.0 * tmpTempError;

            tmpFlowError := flowSP - flowPV;
            tmpTrialValve := accF + 0.5 * tmpFlowError * scanSeconds;
            valveCommand := LIMIT(0.0, 2.0 * tmpFlowError + tmpTrialValve, 100.0);
            accF := valveCommand - 2.0 * tmpFlowError;
        ELSE
            flowSP := manualFlowSP;
            valveCommand := manualValve;
        END_IF;
    ELSE
        IF mode = 0 THEN
            flowSP := manualFlowSP;
            valveCommand := manualValve;
        ELSE
            flowSP := manualFlowSP;
            valveCommand := prevValveCommand;
        END_IF;
    END_IF;
END_IF;

prevMode := mode;
prevResetBtn := resetBtn;
prevNormalMode := normalMode;
prevFlowSP := flowSP;
prevValveCommand := valveCommand;
prevFlowSetpoint := flowSP;
END_FUNCTION_BLOCK

(* ---- self-hard-07.raw_candidate_04.st ---- *)
FUNCTION_BLOCK FB
VAR_INPUT
    mode            : INT;
    resetBtn        : BOOL;
    scanSeconds     : REAL;
    tempSP          : REAL;
    tempPV          : REAL;
    flowPV          : REAL;
    manualFlowSP    : REAL;
    manualValve     : REAL;
END_VAR
VAR_OUTPUT
    flowSP          : REAL;
    valveCommand    : REAL;
    fault           : BOOL;
    normalMode      : BOOL;
END_VAR
VAR
    prevMode            : INT := -1;
    prevResetBtn        : BOOL := FALSE;
    prevNormalMode      : BOOL := FALSE;
    prevFlowSP          : REAL := 0.0;
    prevValveCommand    : REAL := 0.0;
END_VAR
VAR_TEMP
    tmpRisingReset      : BOOL;
    tmpModeChanged      : BOOL;
    tmpTempError        : REAL;
    tmpFlowError        : REAL;
    tmpTrialFlow        : REAL;
    tmpTrialValve       : REAL;
END_VAR
(* ENGINEERING_CONTRACT
 * | Output/State     | Activation          | Retention/Hold         | Explicit Reset   | Same-Scan Priority | Units/Boundaries    |
 * |------------------|---------------------|------------------------|------------------|--------------------|---------------------|
 * | flowSP           | mode=2: cascaded PI | mode=2: hold prev; 0/1: hold prev | reset/fault: follow manualFlowSP | fault/reset > PI calc | 0..50 t/h, KpT=1.0, KiT=0.2/s |
 * | valveCommand     | mode>=1: cascaded PI| mode=1/2: hold prev; 0: follow manual | reset/fault: follow manualValve | fault/reset > PI calc | 0..100 %, KpF=2.0, KiF=0.5/s |
 * | fault            | mode∉{0,1,2} OR scanSeconds∉(0,10] | HOLD until mode/scanSeconds valid | resetBtn↑: cleared | evaluated before reset logic | Boolean |
 * | normalMode       | prevNormalMode AND mode=prevMode AND !fault AND !rising(resetBtn) | mode change: FALSE until re-stabilized | resetBtn↑: FALSE | - | Boolean |
 * | accT (internal)  | mode=2 AND normalMode: back-calc from limited flowSP | mode≠2: retain | reset: 0.0 | PI calc > limit | t/h |
 * | accF (internal)  | mode≥1 AND normalMode: back-calc from limited valveCommand | mode<1: retain | reset: 0.0 | PI calc > limit | % |
 * PUB001: mode ∈ {0,1,2} required for normal; PUB002: scanSeconds ∈ (0,10] required
 * PUB003: resetBtn rising edge triggers re-initialization; PUB004:按住不放不重复动作
 * PUB005: mode switch bumpless: mode=2 holds both, mode=0/1 holds valve; PUB006: PI anti-windup by back-calculation
 * PUB007: first scan outputs initialized to manual values; PUB008: normalMode when stable non-fault non-reset
 *)

(* CONTRACT_RULES [] *)

tmpRisingReset := resetBtn AND NOT prevResetBtn;
tmpModeChanged := (mode <> prevMode);

fault := (mode < 0) OR (mode > 2) OR (scanSeconds <= 0.0) OR (scanSeconds > 10.0);

IF tmpRisingReset THEN
    fault := FALSE;
    normalMode := FALSE;
    accT := 0.0;
    accF := 0.0;
    flowSP := manualFlowSP;
    valveCommand := manualValve;
    prevResetBtn := TRUE;
    prevNormalMode := FALSE;
    prevMode := mode;
    RETURN;
END_IF;

IF prevMode = -1 THEN
    normalMode := FALSE;
    flowSP := manualFlowSP;
    valveCommand := manualValve;
    prevMode := mode;
    prevResetBtn := resetBtn;
    prevNormalMode := TRUE;
    RETURN;
END_IF;

IF tmpModeChanged AND NOT fault THEN
    normalMode := FALSE;
    prevNormalMode := FALSE;
    IF mode = 2 THEN
        flowSP := prevFlowSP;
        valveCommand := prevValveCommand;
    ELSE
        flowSP := manualFlowSP;
        valveCommand := prevValveCommand;
    END_IF;
ELSE
    normalMode := prevNormalMode AND (mode = prevMode) AND NOT fault AND NOT tmpRisingReset;
    IF normalMode THEN
        tmpTempError := tempSP - tempPV;
        tmpTrialFlow := accT + 0.2 * tmpTempError * scanSeconds;
        flowSP := LIMIT(0.0, 1.0 * tmpTempError + tmpTrialFlow, 50.0);
        accT := flowSP - 1.0 * tmpTempError;

        tmpFlowError := flowSP - flowPV;
        tmpTrialValve := accF + 0.5 * tmpFlowError * scanSeconds;
        valveCommand := LIMIT(0.0, 2.0 * tmpFlowError + tmpTrialValve, 100.0);
        accF := valveCommand - 2.0 * tmpFlowError;
    END_IF;
END_IF;

prevMode := mode;
prevResetBtn := resetBtn;
prevNormalMode := normalMode;
prevFlowSP := flowSP;
prevValveCommand := valveCommand;
END_FUNCTION_BLOCK

(* ---- self-medium-01.candidate_01.st ---- *)
TYPE ST_Recipe :
STRUCT
    recipeID    : INT;
    totalRatio  : REAL;
    temperature : REAL;
END_STRUCT
END_TYPE;

FUNCTION_BLOCK FB
VAR_INPUT
    recipe   : ARRAY[1..8] OF ST_Recipe;
    selSlot  : INT;
    loadCmd  : BOOL;
    running  : BOOL;
END_VAR
VAR_OUTPUT
    valid    : BOOL;
    loadedID : INT;
END_VAR
VAR
    tmp_prevLoadCmd : BOOL := FALSE;
    tmp_loadRising  : BOOL := FALSE;
    tmp_prevRunning : BOOL := FALSE;
    tmp_prevLoadedID : INT := 0;
    tmp_prevValid   : BOOL := FALSE;
END_VAR

(* ENGINEERING_CONTRACT
 * +----------------------------------------------------+-------------------------------+---------------------------+---------------------------+----------------+
 * | Output/State Group | Activation | Retention/Hold  | Explicit Reset/Deactivation  | Same-Scan Priority        | Units/Boundaries |
 * +--------------------+------------+-----------------+-------------------------------+---------------------------+------------------+
 * | valid              | rising(loadCmd) & !running | Hold across scans unless reset | !running & rising(loadCmd)| Same scan as loadedID | BOOL |
 * | loadedID           | rising(loadCmd) & !running | Hold when running or idle      | !running & rising(loadCmd)| Same scan as valid     | INT[0..recipeID]|
 * | tmp_loadRising     | loadCmd & !tmp_prevLoadCmd | Cleared each scan              | N/A (internal edge detect)| N/A               | BOOL |
 * | tmp_prevLoadCmd    | copy loadCmd each scan      | N/A                            | N/A                       | N/A               | BOOL |
 * | tmp_prevRunning    | copy running each scan      | N/A                            | N/A                       | N/A               | BOOL |
 * +--------------------+------------+-----------------+-------------------------------+---------------------------+------------------+
 *
 * PUB001 (loadCmd rising edge): Only activates on transition FALSE->TRUE
 * PUB002 (selSlot 1..8): Out-of-bounds treated as invalid, no array access
 * PUB003 (validation rules): totalRatio[99.0,101.0], temperature[30.0,180.0], recipeID<>0
 * PUB004 (running=TRUE): Blocks load, preserves loadedID/valid
 * PUB005 (loadedID update): valid->recipe[selSlot].recipeID, invalid->0
 * PUB006 (valid output): TRUE when all 3 conditions met
 * PUB007 (no edge repeat): Rising edge only, not level-sensitive
 *
 * CONTRACT_RULES [{"kind":"hold_until_reset","output":"valid","set_input":"loadCmd","reset_input":null},{"kind":"hold_until_reset","output":"loadedID","set_input":"loadCmd","reset_input":null}]
 *)
tmp_loadRising := loadCmd AND NOT tmp_prevLoadCmd;

IF tmp_prevRunning AND running THEN
    valid := tmp_prevValid;
    loadedID := tmp_prevLoadedID;
ELSIF running THEN
    valid := tmp_prevValid;
    loadedID := tmp_prevLoadedID;
ELSIF tmp_loadRising THEN
    IF (selSlot < 1) OR (selSlot > 8) THEN
        valid := FALSE;
        loadedID := 0;
    ELSIF recipe[selSlot].recipeID = 0 THEN
        valid := FALSE;
        loadedID := 0;
    ELSIF (recipe[selSlot].totalRatio < 99.0) OR (recipe[selSlot].totalRatio > 101.0) THEN
        valid := FALSE;
        loadedID := 0;
    ELSIF (recipe[selSlot].temperature < 30.0) OR (recipe[selSlot].temperature > 180.0) THEN
        valid := FALSE;
        loadedID := 0;
    ELSE
        valid := TRUE;
        loadedID := recipe[selSlot].recipeID;
    END_IF;
ELSE
    valid := tmp_prevValid;
    loadedID := tmp_prevLoadedID;
END_IF;

tmp_prevLoadCmd := loadCmd;
tmp_prevRunning := running;
tmp_prevLoadedID := loadedID;
tmp_prevValid := valid;

END_FUNCTION_BLOCK

(* ---- self-medium-01.raw_candidate_01.st ---- *)
TYPE ST_Recipe :
STRUCT
    recipeID    : INT;
    totalRatio  : REAL;
    temperature : REAL;
END_STRUCT
END_TYPE

FUNCTION_BLOCK FB
VAR_INPUT
    recipe   : ARRAY[1..8] OF ST_Recipe;
    selSlot  : INT;
    loadCmd  : BOOL;
    running  : BOOL;
END_VAR
VAR_OUTPUT
    valid    : BOOL;
    loadedID : INT;
END_VAR
VAR
    tmp_prevLoadCmd : BOOL := FALSE;
    tmp_loadRising  : BOOL := FALSE;
    tmp_prevRunning : BOOL := FALSE;
    tmp_prevLoadedID : INT := 0;
    tmp_prevValid   : BOOL := FALSE;
END_VAR

(* ENGINEERING_CONTRACT
 * +----------------------------------------------------+-------------------------------+---------------------------+---------------------------+----------------+
 * | Output/State Group | Activation | Retention/Hold  | Explicit Reset/Deactivation  | Same-Scan Priority        | Units/Boundaries |
 * +--------------------+------------+-----------------+-------------------------------+---------------------------+------------------+
 * | valid              | rising(loadCmd) & !running | Hold across scans unless reset | !running & rising(loadCmd)| Same scan as loadedID | BOOL |
 * | loadedID           | rising(loadCmd) & !running | Hold when running or idle      | !running & rising(loadCmd)| Same scan as valid     | INT[0..recipeID]|
 * | tmp_loadRising     | loadCmd & !tmp_prevLoadCmd | Cleared each scan              | N/A (internal edge detect)| N/A               | BOOL |
 * | tmp_prevLoadCmd    | copy loadCmd each scan      | N/A                            | N/A                       | N/A               | BOOL |
 * | tmp_prevRunning    | copy running each scan      | N/A                            | N/A                       | N/A               | BOOL |
 * +--------------------+------------+-----------------+-------------------------------+---------------------------+------------------+
 *
 * PUB001 (loadCmd rising edge): Only activates on transition FALSE->TRUE
 * PUB002 (selSlot 1..8): Out-of-bounds treated as invalid, no array access
 * PUB003 (validation rules): totalRatio[99.0,101.0], temperature[30.0,180.0], recipeID<>0
 * PUB004 (running=TRUE): Blocks load, preserves loadedID/valid
 * PUB005 (loadedID update): valid->recipe[selSlot].recipeID, invalid->0
 * PUB006 (valid output): TRUE when all 3 conditions met
 * PUB007 (no edge repeat): Rising edge only, not level-sensitive
 *
 * CONTRACT_RULES [{"kind":"hold_until_reset","output":"valid","set_input":"loadCmd","reset_input":null},{"kind":"hold_until_reset","output":"loadedID","set_input":"loadCmd","reset_input":null}]
 *)
tmp_loadRising := loadCmd AND NOT tmp_prevLoadCmd;

IF tmp_prevRunning AND running THEN
    valid := tmp_prevValid;
    loadedID := tmp_prevLoadedID;
ELSIF running THEN
    valid := tmp_prevValid;
    loadedID := tmp_prevLoadedID;
ELSIF tmp_loadRising THEN
    IF (selSlot < 1) OR (selSlot > 8) THEN
        valid := FALSE;
        loadedID := 0;
    ELSIF recipe[selSlot].recipeID = 0 THEN
        valid := FALSE;
        loadedID := 0;
    ELSIF (recipe[selSlot].totalRatio < 99.0) OR (recipe[selSlot].totalRatio > 101.0) THEN
        valid := FALSE;
        loadedID := 0;
    ELSIF (recipe[selSlot].temperature < 30.0) OR (recipe[selSlot].temperature > 180.0) THEN
        valid := FALSE;
        loadedID := 0;
    ELSE
        valid := TRUE;
        loadedID := recipe[selSlot].recipeID;
    END_IF;
ELSE
    valid := tmp_prevValid;
    loadedID := tmp_prevLoadedID;
END_IF;

tmp_prevLoadCmd := loadCmd;
tmp_prevRunning := running;
tmp_prevLoadedID := loadedID;
tmp_prevValid := valid;

END_FUNCTION_BLOCK

(* ---- self-medium-02.candidate_01.st ---- *)
FUNCTION_BLOCK FB
VAR_INPUT
    enable  : BOOL;
    rawValue : REAL;
END_VAR

VAR_OUTPUT
    filteredValue : REAL;
    windowFull    : BOOL;
    sampleCount   : INT;
END_VAR

VAR
    buffer     : ARRAY[0..7] OF REAL;
    writeIndex : INT := 0;
    tmp_sum    : REAL;
    tmp_i      : INT;
END_VAR

(*
ENGINEERING_CONTRACT
====================
State retention: filteredValue holds last computed average when disabled; cleared only on re-enable with fresh buffer.
Activation:     sampleCount increments per scan (0→8 max), windowFull TRUE when count=8, stays TRUE until enable=FALSE.
Explicit reset: enable=FALSE clears sampleCount and windowFull in same scan; filteredValue preserved.
Same-scan priority: All outputs updated before function returns.
Units/boundaries: sampleCount ∈ [0,8], buffer size = 8 REAL slots, circular overwrite when full.

Contract Rules: []
*)

IF enable THEN
    // Buffer not yet full: grow window
    IF sampleCount < 8 THEN
        buffer[writeIndex] := rawValue;
        sampleCount := sampleCount + 1;
        writeIndex := (writeIndex + 1) MOD 8;
    ELSE
        // Buffer full: overwrite oldest via circular index
        buffer[writeIndex] := rawValue;
        writeIndex := (writeIndex + 1) MOD 8;
    END_IF;
ELSE
    // Disable: clear count and full flag, retain filteredValue
    sampleCount := 0;
    windowFull  := FALSE;
END_IF;

// Compute filteredValue from valid samples only
tmp_sum := 0.0;
FOR tmp_i := 0 TO sampleCount - 1 DO
    tmp_sum := tmp_sum + buffer[tmp_i];
END_FOR;

IF sampleCount > 0 THEN
    filteredValue := tmp_sum / TO_REAL(sampleCount);
    windowFull := (sampleCount = 8);
ELSE
    filteredValue := 0.0;
END_IF;

END_FUNCTION_BLOCK

(* ---- self-medium-02.candidate_02.st ---- *)
FUNCTION_BLOCK FB
VAR_INPUT
    enable   : BOOL;
    rawValue : REAL;
END_VAR

VAR_OUTPUT
    filteredValue : REAL;
    windowFull    : BOOL;
    sampleCount   : INT;
END_VAR

VAR
    buffer      : ARRAY[0..7] OF REAL;
    writeIndex  : INT := 0;
    bufferValid : BOOL := FALSE;
    tmp_sum     : REAL;
    tmp_i       : INT;
END_VAR

(*
ENGINEERING_CONTRACT
====================
State retention: filteredValue holds last computed average when disabled; cleared only on re-enable with fresh buffer.
Activation:     sampleCount increments per scan (0→8 max), windowFull TRUE when count=8, stays TRUE until enable=FALSE.
Explicit reset: enable=FALSE clears sampleCount and windowFull in same scan; filteredValue preserved.
Same-scan priority: All outputs updated before function returns.
Units/boundaries: sampleCount ∈ [0,8], buffer size = 8 REAL slots, circular overwrite when full.

Contract Rules: []
*)

IF enable THEN
    // First sample after disable: invalidate old buffer
    IF NOT bufferValid THEN
        writeIndex  := 0;
        sampleCount := 0;
    END_IF;
    bufferValid := TRUE;

    // Buffer not yet full: grow window
    IF sampleCount < 8 THEN
        buffer[writeIndex] := rawValue;
        sampleCount := sampleCount + 1;
        writeIndex := (writeIndex + 1) MOD 8;
    ELSE
        // Buffer full: overwrite oldest via circular index
        buffer[writeIndex] := rawValue;
        writeIndex := (writeIndex + 1) MOD 8;
    END_IF;

    // Compute filteredValue from valid samples only
    tmp_sum := 0.0;
    FOR tmp_i := 0 TO sampleCount - 1 DO
        tmp_sum := tmp_sum + buffer[tmp_i];
    END_FOR;
    filteredValue := tmp_sum / TO_REAL(sampleCount);
    windowFull := (sampleCount = 8);
ELSE
    // Disable: clear count and full flag, retain filteredValue and buffer
    bufferValid := FALSE;
    sampleCount := 0;
    windowFull  := FALSE;
END_IF;

END_FUNCTION_BLOCK

(* ---- self-medium-02.raw_candidate_01.st ---- *)
FUNCTION_BLOCK FB
VAR_INPUT
    enable  : BOOL;
    rawValue : REAL;
END_VAR

VAR_OUTPUT
    filteredValue : REAL;
    windowFull    : BOOL;
    sampleCount   : INT;
END_VAR

VAR
    buffer     : ARRAY[0..7] OF REAL;
    writeIndex : INT := 0;
    tmp_sum    : REAL;
    tmp_i      : INT;
END_VAR

(*
ENGINEERING_CONTRACT
====================
State retention: filteredValue holds last computed average when disabled; cleared only on re-enable with fresh buffer.
Activation:     sampleCount increments per scan (0→8 max), windowFull TRUE when count=8, stays TRUE until enable=FALSE.
Explicit reset: enable=FALSE clears sampleCount and windowFull in same scan; filteredValue preserved.
Same-scan priority: All outputs updated before function returns.
Units/boundaries: sampleCount ∈ [0,8], buffer size = 8 REAL slots, circular overwrite when full.

Contract Rules: []
*)

IF enable THEN
    // Buffer not yet full: grow window
    IF sampleCount < 8 THEN
        buffer[writeIndex] := rawValue;
        sampleCount := sampleCount + 1;
        writeIndex := (writeIndex + 1) MOD 8;
    ELSE
        // Buffer full: overwrite oldest via circular index
        buffer[writeIndex] := rawValue;
        writeIndex := (writeIndex + 1) MOD 8;
    END_IF;
ELSE
    // Disable: clear count and full flag, retain filteredValue
    sampleCount := 0;
    windowFull  := FALSE;
END_IF;

// Compute filteredValue from valid samples only
tmp_sum := 0.0;
FOR tmp_i := 0 TO sampleCount - 1 DO
    tmp_sum := tmp_sum + buffer[tmp_i];
END_FOR;

IF sampleCount > 0 THEN
    filteredValue := tmp_sum / TO_REAL(sampleCount);
    windowFull := (sampleCount = 8);
ELSE
    filteredValue := 0.0;
END_IF;

END_FUNCTION_BLOCK

(* ---- self-medium-02.raw_candidate_02.st ---- *)
FUNCTION_BLOCK FB
VAR_INPUT
    enable   : BOOL;
    rawValue : REAL;
END_VAR

VAR_OUTPUT
    filteredValue : REAL;
    windowFull    : BOOL;
    sampleCount   : INT;
END_VAR

VAR
    buffer      : ARRAY[0..7] OF REAL;
    writeIndex  : INT := 0;
    bufferValid : BOOL := FALSE;
    tmp_sum     : REAL;
    tmp_i       : INT;
END_VAR

(*
ENGINEERING_CONTRACT
====================
State retention: filteredValue holds last computed average when disabled; cleared only on re-enable with fresh buffer.
Activation:     sampleCount increments per scan (0→8 max), windowFull TRUE when count=8, stays TRUE until enable=FALSE.
Explicit reset: enable=FALSE clears sampleCount and windowFull in same scan; filteredValue preserved.
Same-scan priority: All outputs updated before function returns.
Units/boundaries: sampleCount ∈ [0,8], buffer size = 8 REAL slots, circular overwrite when full.

Contract Rules: []
*)

IF enable THEN
    // First sample after disable: invalidate old buffer
    IF NOT bufferValid THEN
        writeIndex  := 0;
        sampleCount := 0;
    END_IF;
    bufferValid := TRUE;

    // Buffer not yet full: grow window
    IF sampleCount < 8 THEN
        buffer[writeIndex] := rawValue;
        sampleCount := sampleCount + 1;
        writeIndex := (writeIndex + 1) MOD 8;
    ELSE
        // Buffer full: overwrite oldest via circular index
        buffer[writeIndex] := rawValue;
        writeIndex := (writeIndex + 1) MOD 8;
    END_IF;

    // Compute filteredValue from valid samples only
    tmp_sum := 0.0;
    FOR tmp_i := 0 TO sampleCount - 1 DO
        tmp_sum := tmp_sum + buffer[tmp_i];
    END_FOR;
    filteredValue := tmp_sum / TO_REAL(sampleCount);
    windowFull := (sampleCount = 8);
ELSE
    // Disable: clear count and full flag, retain filteredValue and buffer
    bufferValid := FALSE;
    sampleCount := 0;
    windowFull  := FALSE;
END_IF;

END_FUNCTION_BLOCK

(* ---- self-medium-03.candidate_01.st ---- *)
FUNCTION_BLOCK FB
VAR_INPUT
    openBtn    : BOOL;
    closeBtn   : BOOL;
    openLimit  : BOOL;
    closeLimit : BOOL;
    obstacle   : BOOL;
END_VAR
VAR_OUTPUT
    motorUp    : BOOL;
    motorDown  : BOOL;
    errorFlag  : BOOL;
END_VAR
VAR
    state       : EState := IDLE;
    prev_openBtn   : BOOL := FALSE;
    prev_closeBtn  : BOOL := FALSE;
    prev_obstacle  : BOOL := FALSE;
    openRTrig      : R_TRIG;
    closeRTrig     : R_TRIG;
    dualRTrig      : R_TRIG;
END_VAR

(*
ENGINEERING_CONTRACT
===================
| Output/State | Activation          | Retention          | Reset/Deactivation        | Scan Priority | Units      |
|--------------|---------------------|--------------------|---------------------------|---------------|------------|
| motorUp      | IDLE+rising(openBtn)| Running continues  | obstacle/closeLimit/FAULT | Same-scan     | BOOL       |
| motorDown    | IDLE+rising(closeBtn)| Running continues | obstacle/openLimit/FAULT  | Same-scan     | BOOL       |
| errorFlag    | Any state+obstacle  | Latched in FAULT   | No obstacle+dualBtn rising| Highest      | BOOL       |
| state=FAULT  | Any state+obstacle  | Until dualBtn reset| No obstacle+dualBtn rising| Highest      | EState     |
| state=IDLE   | Power-on/limit/reset| Until openBtn/closeBtn rising | -                  | Default     | EState     |
PUB001: power-on IDLE
PUB002: init FALSE
PUB003: no obstacle IDLE start rules (openBtn edge, closeBtn=FALSE, not openLimit)
PUB004: no obstacle close start rules (closeBtn edge, openBtn=FALSE, not closeLimit)
PUB006: no dual-btn start
PUB007: same-scan motor command on start
PUB008: button release ignored during movement
PUB009: direction buttons ignored during movement
PUB010: limit stop same-scan
PUB011: opposite limit does not affect
PUB012: mutual exclusion always
PUB013: obstacle immediate both-stop + FAULT
PUB014: FAULT priority over limits/movement/reset
PUB017: errorFlag latched
PUB018: FAULT stop motors
PUB019: reset requires no obstacle + dualBtn from not-both to both
PUB020: cannot reset during obstacle
PUB021: cannot auto-reset on obstacle clear
PUB022: reset → IDLE
PUB023: reset same-scan both motors stop
PUB024: post-reset follow rule 1
*)
BEGIN
    openRTrig(CLK := openBtn);
    closeRTrig(CLK := closeBtn);
    dualRTrig(CLK := openBtn AND closeBtn);

    (* Priority 1: Obstacle → immediate stop + FAULT *)
    IF obstacle THEN
        motorUp   := FALSE;
        motorDown := FALSE;
        state     := FAULT;
        errorFlag := TRUE;
    ELSE
        CASE state OF
            IDLE:
                motorUp   := FALSE;
                motorDown := FALSE;

                (* Start opening *)
                IF openRTrig.Q AND NOT closeBtn AND NOT openLimit THEN
                    motorUp := TRUE;
                    state   := OPENING;
                (* Start closing *)
                ELSIF closeRTrig.Q AND NOT openBtn AND NOT closeLimit THEN
                    motorDown := TRUE;
                    state     := CLOSING;
                END_IF;

            OPENING:
                motorUp   := TRUE;
                motorDown := FALSE;
                IF openLimit THEN
                    motorUp := FALSE;
                    state   := IDLE;
                END_IF;

            CLOSING:
                motorUp   := FALSE;
                motorDown := TRUE;
                IF closeLimit THEN
                    motorDown := FALSE;
                    state     := IDLE;
                END_IF;

            FAULT:
                motorUp   := FALSE;
                motorDown := FALSE;
                IF dualRTrig.Q THEN
                    errorFlag := FALSE;
                    state     := IDLE;
                END_IF;
        END_CASE;
    END_IF;

    prev_openBtn  := openBtn;
    prev_closeBtn := closeBtn;
    prev_obstacle := obstacle;
END_FUNCTION_BLOCK

TYPE EState : (
    IDLE    := 0,
    OPENING := 1,
    CLOSING := 2,
    FAULT   := 3
) END_TYPE;
END_TYPE;

(* CONTRACT_RULES [] *)

(* ---- self-medium-03.candidate_02.st ---- *)
FUNCTION_BLOCK FB
VAR_INPUT
    openBtn    : BOOL;
    closeBtn   : BOOL;
    openLimit  : BOOL;
    closeLimit : BOOL;
    obstacle   : BOOL;
END_VAR
VAR_OUTPUT
    motorUp    : BOOL;
    motorDown  : BOOL;
    errorFlag  : BOOL;
END_VAR
VAR
    state         : EState := IDLE;
    prev_openBtn  : BOOL := FALSE;
    prev_closeBtn : BOOL := FALSE;
    openRTrig     : R_TRIG;
    closeRTrig    : R_TRIG;
    dualRTrig     : R_TRIG;
END_VAR

(*
ENGINEERING_CONTRACT
===================
| Output/State | Activation          | Retention          | Reset/Deactivation        | Scan Priority | Units      |
|--------------|---------------------|--------------------|---------------------------|---------------|------------|
| motorUp      | IDLE+rising(openBtn)| Running continues  | obstacle/closeLimit/FAULT | Same-scan     | BOOL       |
| motorDown    | IDLE+rising(closeBtn)| Running continues | obstacle/openLimit/FAULT  | Same-scan     | BOOL       |
| errorFlag    | Any state+obstacle  | Latched in FAULT   | No obstacle+dualBtn rising| Highest      | BOOL       |
| state=FAULT  | Any state+obstacle  | Until dualBtn reset| No obstacle+dualBtn rising| Highest      | EState     |
| state=IDLE   | Power-on/limit/reset| Until openBtn/closeBtn rising | -                  | Default     | EState     |
PUB001: power-on IDLE
PUB002: init FALSE
PUB003: no obstacle IDLE start rules (openBtn edge, closeBtn=FALSE, not openLimit)
PUB004: no obstacle close start rules (closeBtn edge, openBtn=FALSE, not closeLimit)
PUB006: no dual-btn start
PUB007: same-scan motor command on start
PUB008: button release ignored during movement
PUB009: direction buttons ignored during movement
PUB010: limit stop same-scan
PUB011: opposite limit does not affect
PUB012: mutual exclusion always
PUB013: obstacle immediate both-stop + FAULT
PUB014: FAULT priority over limits/movement/reset
PUB017: errorFlag latched
PUB018: FAULT stop motors
PUB019: reset requires no obstacle + dualBtn from not-both to both
PUB020: cannot reset during obstacle
PUB021: cannot auto-reset on obstacle clear
PUB022: reset → IDLE
PUB023: reset same-scan both motors stop
PUB024: post-reset follow rule 1
*)
BEGIN
    openRTrig(CLK := openBtn);
    closeRTrig(CLK := closeBtn);
    dualRTrig(CLK := openBtn AND closeBtn);

    (* Priority 1: Obstacle → immediate stop + FAULT *)
    IF obstacle THEN
        motorUp   := FALSE;
        motorDown := FALSE;
        state     := FAULT;
        errorFlag := TRUE;
    ELSE
        CASE state OF
            IDLE:
                motorUp   := FALSE;
                motorDown := FALSE;

                (* Start opening *)
                IF openRTrig.Q AND NOT closeBtn AND NOT openLimit THEN
                    motorUp := TRUE;
                    state   := OPENING;
                (* Start closing *)
                ELSIF closeRTrig.Q AND NOT openBtn AND NOT closeLimit THEN
                    motorDown := TRUE;
                    state     := CLOSING;
                END_IF;

            OPENING:
                motorUp   := TRUE;
                motorDown := FALSE;
                IF openLimit THEN
                    motorUp := FALSE;
                    state   := IDLE;
                END_IF;

            CLOSING:
                motorUp   := FALSE;
                motorDown := TRUE;
                IF closeLimit THEN
                    motorDown := FALSE;
                    state     := IDLE;
                END_IF;

            FAULT:
                motorUp   := FALSE;
                motorDown := FALSE;
                IF dualRTrig.Q THEN
                    errorFlag := FALSE;
                    state     := IDLE;
                END_IF;
        END_CASE;
    END_IF;

    prev_openBtn  := openBtn;
    prev_closeBtn := closeBtn;
END_FUNCTION_BLOCK

TYPE EState : (
    IDLE    := 0,
    OPENING := 1,
    CLOSING := 2,
    FAULT   := 3
) END_TYPE;

(* CONTRACT_RULES [] *)

(* ---- self-medium-03.candidate_03.st ---- *)
TYPE EState : (
    IDLE    := 0,
    OPENING := 1,
    CLOSING := 2,
    FAULT   := 3
) END_TYPE;

FUNCTION_BLOCK FB
VAR_INPUT
    openBtn    : BOOL;
    closeBtn   : BOOL;
    openLimit  : BOOL;
    closeLimit : BOOL;
    obstacle   : BOOL;
END_VAR
VAR_OUTPUT
    motorUp    : BOOL;
    motorDown  : BOOL;
    errorFlag  : BOOL;
END_VAR
VAR
    state       : EState := IDLE;
    prev_openBtn   : BOOL := FALSE;
    prev_closeBtn  : BOOL := FALSE;
    prev_obstacle  : BOOL := FALSE;
    openRTrig      : R_TRIG;
    closeRTrig     : R_TRIG;
    dualRTrig      : R_TRIG;
END_VAR

(*
ENGINEERING_CONTRACT
===================
| Output/State | Activation          | Retention          | Reset/Deactivation        | Scan Priority | Units      |
|--------------|---------------------|--------------------|---------------------------|---------------|------------|
| motorUp      | IDLE+rising(openBtn)| Running continues  | obstacle/closeLimit/FAULT | Same-scan     | BOOL       |
| motorDown    | IDLE+rising(closeBtn)| Running continues | obstacle/openLimit/FAULT  | Same-scan     | BOOL       |
| errorFlag    | Any state+obstacle  | Latched in FAULT   | No obstacle+dualBtn rising| Highest      | BOOL       |
| state=FAULT  | Any state+obstacle  | Until dualBtn reset| No obstacle+dualBtn rising| Highest      | EState     |
| state=IDLE   | Power-on/limit/reset| Until openBtn/closeBtn rising | -                  | Default     | EState     |
PUB001: power-on IDLE
PUB002: init FALSE
PUB003: no obstacle IDLE start rules (openBtn edge, closeBtn=FALSE, not openLimit)
PUB004: no obstacle close start rules (closeBtn edge, openBtn=FALSE, not closeLimit)
PUB006: no dual-btn start
PUB007: same-scan motor command on start
PUB008: button release ignored during movement
PUB009: direction buttons ignored during movement
PUB010: limit stop same-scan
PUB011: opposite limit does not affect
PUB012: mutual exclusion always
PUB013: obstacle immediate both-stop + FAULT
PUB014: FAULT priority over limits/movement/reset
PUB017: errorFlag latched
PUB018: FAULT stop motors
PUB019: reset requires no obstacle + dualBtn from not-both to both
PUB020: cannot reset during obstacle
PUB021: cannot auto-reset on obstacle clear
PUB022: reset → IDLE
PUB023: reset same-scan both motors stop
PUB024: post-reset follow rule 1
*)
BEGIN
    openRTrig(CLK := openBtn);
    closeRTrig(CLK := closeBtn);
    dualRTrig(CLK := openBtn AND closeBtn);

    (* Priority 1: Obstacle → immediate stop + FAULT *)
    IF obstacle THEN
        motorUp   := FALSE;
        motorDown := FALSE;
        state     := FAULT;
        errorFlag := TRUE;
    ELSE
        CASE state OF
            IDLE:
                motorUp   := FALSE;
                motorDown := FALSE;

                (* Start opening *)
                IF openRTrig.Q AND NOT closeBtn AND NOT openLimit THEN
                    motorUp := TRUE;
                    state   := OPENING;
                (* Start closing *)
                ELSIF closeRTrig.Q AND NOT openBtn AND NOT closeLimit THEN
                    motorDown := TRUE;
                    state     := CLOSING;
                END_IF;

            OPENING:
                motorUp   := TRUE;
                motorDown := FALSE;
                IF openLimit THEN
                    motorUp := FALSE;
                    state   := IDLE;
                END_IF;

            CLOSING:
                motorUp   := FALSE;
                motorDown := TRUE;
                IF closeLimit THEN
                    motorDown := FALSE;
                    state     := IDLE;
                END_IF;

            FAULT:
                motorUp   := FALSE;
                motorDown := FALSE;
                IF dualRTrig.Q THEN
                    errorFlag := FALSE;
                    state     := IDLE;
                END_IF;
        END_CASE;
    END_IF;

    prev_openBtn  := openBtn;
    prev_closeBtn := closeBtn;
    prev_obstacle := obstacle;
END_FUNCTION_BLOCK

(* CONTRACT_RULES [] *)

(* ---- self-medium-03.candidate_04.st ---- *)
TYPE EState :
    (
        IDLE    := 0,
        OPENING := 1,
        CLOSING := 2,
        FAULT   := 3
    )
END_TYPE;

FUNCTION_BLOCK FB
VAR_INPUT
    openBtn    : BOOL;
    closeBtn   : BOOL;
    openLimit  : BOOL;
    closeLimit : BOOL;
    obstacle   : BOOL;
END_VAR
VAR_OUTPUT
    motorUp    : BOOL;
    motorDown  : BOOL;
    errorFlag  : BOOL;
END_VAR
VAR
    state          : EState := IDLE;
    prev_openBtn   : BOOL := FALSE;
    prev_closeBtn  : BOOL := FALSE;
    prev_obstacle  : BOOL := FALSE;
    openRTrig      : R_TRIG;
    closeRTrig     : R_TRIG;
    dualRTrig      : R_TRIG;
END_VAR

(*
ENGINEERING_CONTRACT
===================
| Output/State | Activation           | Retention           | Reset/Deactivation              | Scan Priority | Units   |
|--------------|----------------------|---------------------|----------------------------------|---------------|---------|
| motorUp      | IDLE+rising(openBtn) | Running continues   | obstacle/openLimit/FAULT         | Same-scan     | BOOL    |
| motorDown    | IDLE+rising(closeBtn)| Running continues   | obstacle/closeLimit/FAULT        | Same-scan     | BOOL    |
| errorFlag    | Any state+obstacle   | Latched in FAULT    | No obstacle+dualBtn rising edge  | Highest       | BOOL    |
| state=FAULT  | Any state+obstacle   | Until dualBtn reset | No obstacle+dualBtn rising edge  | Highest       | EState  |
| state=IDLE   | Power-on/limit/reset | Until rising edge   | -                                | Default       | EState  |
PUB001: power-on IDLE
PUB002: init FALSE
PUB003-005: no obstacle IDLE start (openBtn rising, closeBtn=FALSE, not openLimit)
PUB006: dual-btn does not start
PUB007: motor command same-scan on start
PUB008-009: button release / direction buttons ignored during movement
PUB010-011: limit stop same-scan, opposite limit irrelevant
PUB012: mutual exclusion always
PUB013-014: obstacle → both stop + FAULT (highest priority)
PUB017-018: errorFlag latched, motors stopped in FAULT
PUB019-021: reset requires no obstacle + dualBtn from not-both to both
PUB022-024: reset → IDLE, same-scan stop, then follow rule 1
*)

BEGIN
    openRTrig(CLK := openBtn);
    closeRTrig(CLK := closeBtn);
    dualRTrig(CLK := openBtn AND closeBtn);

    (* Priority 1: Obstacle → immediate both-stop + FAULT *)
    IF obstacle THEN
        motorUp   := FALSE;
        motorDown := FALSE;
        state     := FAULT;
        errorFlag := TRUE;
    ELSE
        CASE state OF
            IDLE:
                motorUp   := FALSE;
                motorDown := FALSE;
                (* Start opening: rising edge of openBtn, closeBtn=FALSE, not at openLimit *)
                IF openRTrig.Q AND NOT closeBtn AND NOT openLimit THEN
                    motorUp := TRUE;
                    state   := OPENING;
                (* Start closing: rising edge of closeBtn, openBtn=FALSE, not at closeLimit *)
                ELSIF closeRTrig.Q AND NOT openBtn AND NOT closeLimit THEN
                    motorDown := TRUE;
                    state     := CLOSING;
                END_IF;

            OPENING:
                motorUp   := TRUE;
                motorDown := FALSE;
                IF openLimit THEN
                    motorUp := FALSE;
                    state   := IDLE;
                END_IF;

            CLOSING:
                motorUp   := FALSE;
                motorDown := TRUE;
                IF closeLimit THEN
                    motorDown := FALSE;
                    state     := IDLE;
                END_IF;

            FAULT:
                motorUp   := FALSE;
                motorDown := FALSE;
                IF dualRTrig.Q THEN
                    errorFlag := FALSE;
                    state     := IDLE;
                END_IF;
        END_CASE;
    END_IF;

    prev_openBtn  := openBtn;
    prev_closeBtn := closeBtn;
    prev_obstacle := obstacle;
END_FUNCTION_BLOCK

(* CONTRACT_RULES [] *)

(* ---- self-medium-03.raw_candidate_01.st ---- *)
FUNCTION_BLOCK FB
VAR_INPUT
    openBtn    : BOOL;
    closeBtn   : BOOL;
    openLimit  : BOOL;
    closeLimit : BOOL;
    obstacle   : BOOL;
END_VAR
VAR_OUTPUT
    motorUp    : BOOL;
    motorDown  : BOOL;
    errorFlag  : BOOL;
END_VAR
VAR
    state       : EState := IDLE;
    prev_openBtn   : BOOL := FALSE;
    prev_closeBtn  : BOOL := FALSE;
    prev_obstacle  : BOOL := FALSE;
    openRTrig      : R_TRIG;
    closeRTrig     : R_TRIG;
    dualRTrig      : R_TRIG;
END_VAR

(*
ENGINEERING_CONTRACT
===================
| Output/State | Activation          | Retention          | Reset/Deactivation        | Scan Priority | Units      |
|--------------|---------------------|--------------------|---------------------------|---------------|------------|
| motorUp      | IDLE+rising(openBtn)| Running continues  | obstacle/closeLimit/FAULT | Same-scan     | BOOL       |
| motorDown    | IDLE+rising(closeBtn)| Running continues | obstacle/openLimit/FAULT  | Same-scan     | BOOL       |
| errorFlag    | Any state+obstacle  | Latched in FAULT   | No obstacle+dualBtn rising| Highest      | BOOL       |
| state=FAULT  | Any state+obstacle  | Until dualBtn reset| No obstacle+dualBtn rising| Highest      | EState     |
| state=IDLE   | Power-on/limit/reset| Until openBtn/closeBtn rising | -                  | Default     | EState     |
PUB001: power-on IDLE
PUB002: init FALSE
PUB003: no obstacle IDLE start rules (openBtn edge, closeBtn=FALSE, not openLimit)
PUB004: no obstacle close start rules (closeBtn edge, openBtn=FALSE, not closeLimit)
PUB006: no dual-btn start
PUB007: same-scan motor command on start
PUB008: button release ignored during movement
PUB009: direction buttons ignored during movement
PUB010: limit stop same-scan
PUB011: opposite limit does not affect
PUB012: mutual exclusion always
PUB013: obstacle immediate both-stop + FAULT
PUB014: FAULT priority over limits/movement/reset
PUB017: errorFlag latched
PUB018: FAULT stop motors
PUB019: reset requires no obstacle + dualBtn from not-both to both
PUB020: cannot reset during obstacle
PUB021: cannot auto-reset on obstacle clear
PUB022: reset → IDLE
PUB023: reset same-scan both motors stop
PUB024: post-reset follow rule 1
*)
BEGIN
    openRTrig(CLK := openBtn);
    closeRTrig(CLK := closeBtn);
    dualRTrig(CLK := openBtn AND closeBtn);

    (* Priority 1: Obstacle → immediate stop + FAULT *)
    IF obstacle THEN
        motorUp   := FALSE;
        motorDown := FALSE;
        state     := FAULT;
        errorFlag := TRUE;
    ELSE
        CASE state OF
            IDLE:
                motorUp   := FALSE;
                motorDown := FALSE;

                (* Start opening *)
                IF openRTrig.Q AND NOT closeBtn AND NOT openLimit THEN
                    motorUp := TRUE;
                    state   := OPENING;
                (* Start closing *)
                ELSIF closeRTrig.Q AND NOT openBtn AND NOT closeLimit THEN
                    motorDown := TRUE;
                    state     := CLOSING;
                END_IF

            OPENING:
                motorUp   := TRUE;
                motorDown := FALSE;
                IF openLimit THEN
                    motorUp := FALSE;
                    state   := IDLE;
                END_IF

            CLOSING:
                motorUp   := FALSE;
                motorDown := TRUE;
                IF closeLimit THEN
                    motorDown := FALSE;
                    state     := IDLE;
                END_IF

            FAULT:
                motorUp   := FALSE;
                motorDown := FALSE;
                IF dualRTrig.Q THEN
                    errorFlag := FALSE;
                    state     := IDLE;
                END_IF
        END_CASE
    END_IF

    prev_openBtn  := openBtn;
    prev_closeBtn := closeBtn;
    prev_obstacle := obstacle;
END_FUNCTION_BLOCK

TYPE EState : (
    IDLE    := 0,
    OPENING := 1,
    CLOSING := 2,
    FAULT   := 3
) END_TYPE
END_TYPE

(* CONTRACT_RULES [] *)

(* ---- self-medium-03.raw_candidate_02.st ---- *)
FUNCTION_BLOCK FB
VAR_INPUT
    openBtn    : BOOL;
    closeBtn   : BOOL;
    openLimit  : BOOL;
    closeLimit : BOOL;
    obstacle   : BOOL;
END_VAR
VAR_OUTPUT
    motorUp    : BOOL;
    motorDown  : BOOL;
    errorFlag  : BOOL;
END_VAR
VAR
    state         : EState := IDLE;
    prev_openBtn  : BOOL := FALSE;
    prev_closeBtn : BOOL := FALSE;
    openRTrig     : R_TRIG;
    closeRTrig    : R_TRIG;
    dualRTrig     : R_TRIG;
END_VAR

(*
ENGINEERING_CONTRACT
===================
| Output/State | Activation          | Retention          | Reset/Deactivation        | Scan Priority | Units      |
|--------------|---------------------|--------------------|---------------------------|---------------|------------|
| motorUp      | IDLE+rising(openBtn)| Running continues  | obstacle/closeLimit/FAULT | Same-scan     | BOOL       |
| motorDown    | IDLE+rising(closeBtn)| Running continues | obstacle/openLimit/FAULT  | Same-scan     | BOOL       |
| errorFlag    | Any state+obstacle  | Latched in FAULT   | No obstacle+dualBtn rising| Highest      | BOOL       |
| state=FAULT  | Any state+obstacle  | Until dualBtn reset| No obstacle+dualBtn rising| Highest      | EState     |
| state=IDLE   | Power-on/limit/reset| Until openBtn/closeBtn rising | -                  | Default     | EState     |
PUB001: power-on IDLE
PUB002: init FALSE
PUB003: no obstacle IDLE start rules (openBtn edge, closeBtn=FALSE, not openLimit)
PUB004: no obstacle close start rules (closeBtn edge, openBtn=FALSE, not closeLimit)
PUB006: no dual-btn start
PUB007: same-scan motor command on start
PUB008: button release ignored during movement
PUB009: direction buttons ignored during movement
PUB010: limit stop same-scan
PUB011: opposite limit does not affect
PUB012: mutual exclusion always
PUB013: obstacle immediate both-stop + FAULT
PUB014: FAULT priority over limits/movement/reset
PUB017: errorFlag latched
PUB018: FAULT stop motors
PUB019: reset requires no obstacle + dualBtn from not-both to both
PUB020: cannot reset during obstacle
PUB021: cannot auto-reset on obstacle clear
PUB022: reset → IDLE
PUB023: reset same-scan both motors stop
PUB024: post-reset follow rule 1
*)
BEGIN
    openRTrig(CLK := openBtn);
    closeRTrig(CLK := closeBtn);
    dualRTrig(CLK := openBtn AND closeBtn);

    (* Priority 1: Obstacle → immediate stop + FAULT *)
    IF obstacle THEN
        motorUp   := FALSE;
        motorDown := FALSE;
        state     := FAULT;
        errorFlag := TRUE;
    ELSE
        CASE state OF
            IDLE:
                motorUp   := FALSE;
                motorDown := FALSE;

                (* Start opening *)
                IF openRTrig.Q AND NOT closeBtn AND NOT openLimit THEN
                    motorUp := TRUE;
                    state   := OPENING;
                (* Start closing *)
                ELSIF closeRTrig.Q AND NOT openBtn AND NOT closeLimit THEN
                    motorDown := TRUE;
                    state     := CLOSING;
                END_IF;

            OPENING:
                motorUp   := TRUE;
                motorDown := FALSE;
                IF openLimit THEN
                    motorUp := FALSE;
                    state   := IDLE;
                END_IF;

            CLOSING:
                motorUp   := FALSE;
                motorDown := TRUE;
                IF closeLimit THEN
                    motorDown := FALSE;
                    state     := IDLE;
                END_IF;

            FAULT:
                motorUp   := FALSE;
                motorDown := FALSE;
                IF dualRTrig.Q THEN
                    errorFlag := FALSE;
                    state     := IDLE;
                END_IF;
        END_CASE;
    END_IF;

    prev_openBtn  := openBtn;
    prev_closeBtn := closeBtn;
END_FUNCTION_BLOCK

TYPE EState : (
    IDLE    := 0,
    OPENING := 1,
    CLOSING := 2,
    FAULT   := 3
) END_TYPE;

(* CONTRACT_RULES [] *)

(* ---- self-medium-03.raw_candidate_03.st ---- *)
TYPE EState : (
    IDLE    := 0,
    OPENING := 1,
    CLOSING := 2,
    FAULT   := 3
) END_TYPE;

FUNCTION_BLOCK FB
VAR_INPUT
    openBtn    : BOOL;
    closeBtn   : BOOL;
    openLimit  : BOOL;
    closeLimit : BOOL;
    obstacle   : BOOL;
END_VAR
VAR_OUTPUT
    motorUp    : BOOL;
    motorDown  : BOOL;
    errorFlag  : BOOL;
END_VAR
VAR
    state       : EState := IDLE;
    prev_openBtn   : BOOL := FALSE;
    prev_closeBtn  : BOOL := FALSE;
    prev_obstacle  : BOOL := FALSE;
    openRTrig      : R_TRIG;
    closeRTrig     : R_TRIG;
    dualRTrig      : R_TRIG;
END_VAR

(*
ENGINEERING_CONTRACT
===================
| Output/State | Activation          | Retention          | Reset/Deactivation        | Scan Priority | Units      |
|--------------|---------------------|--------------------|---------------------------|---------------|------------|
| motorUp      | IDLE+rising(openBtn)| Running continues  | obstacle/closeLimit/FAULT | Same-scan     | BOOL       |
| motorDown    | IDLE+rising(closeBtn)| Running continues | obstacle/openLimit/FAULT  | Same-scan     | BOOL       |
| errorFlag    | Any state+obstacle  | Latched in FAULT   | No obstacle+dualBtn rising| Highest      | BOOL       |
| state=FAULT  | Any state+obstacle  | Until dualBtn reset| No obstacle+dualBtn rising| Highest      | EState     |
| state=IDLE   | Power-on/limit/reset| Until openBtn/closeBtn rising | -                  | Default     | EState     |
PUB001: power-on IDLE
PUB002: init FALSE
PUB003: no obstacle IDLE start rules (openBtn edge, closeBtn=FALSE, not openLimit)
PUB004: no obstacle close start rules (closeBtn edge, openBtn=FALSE, not closeLimit)
PUB006: no dual-btn start
PUB007: same-scan motor command on start
PUB008: button release ignored during movement
PUB009: direction buttons ignored during movement
PUB010: limit stop same-scan
PUB011: opposite limit does not affect
PUB012: mutual exclusion always
PUB013: obstacle immediate both-stop + FAULT
PUB014: FAULT priority over limits/movement/reset
PUB017: errorFlag latched
PUB018: FAULT stop motors
PUB019: reset requires no obstacle + dualBtn from not-both to both
PUB020: cannot reset during obstacle
PUB021: cannot auto-reset on obstacle clear
PUB022: reset → IDLE
PUB023: reset same-scan both motors stop
PUB024: post-reset follow rule 1
*)
BEGIN
    openRTrig(CLK := openBtn);
    closeRTrig(CLK := closeBtn);
    dualRTrig(CLK := openBtn AND closeBtn);

    (* Priority 1: Obstacle → immediate stop + FAULT *)
    IF obstacle THEN
        motorUp   := FALSE;
        motorDown := FALSE;
        state     := FAULT;
        errorFlag := TRUE;
    ELSE
        CASE state OF
            IDLE:
                motorUp   := FALSE;
                motorDown := FALSE;

                (* Start opening *)
                IF openRTrig.Q AND NOT closeBtn AND NOT openLimit THEN
                    motorUp := TRUE;
                    state   := OPENING;
                (* Start closing *)
                ELSIF closeRTrig.Q AND NOT openBtn AND NOT closeLimit THEN
                    motorDown := TRUE;
                    state     := CLOSING;
                END_IF;

            OPENING:
                motorUp   := TRUE;
                motorDown := FALSE;
                IF openLimit THEN
                    motorUp := FALSE;
                    state   := IDLE;
                END_IF;

            CLOSING:
                motorUp   := FALSE;
                motorDown := TRUE;
                IF closeLimit THEN
                    motorDown := FALSE;
                    state     := IDLE;
                END_IF;

            FAULT:
                motorUp   := FALSE;
                motorDown := FALSE;
                IF dualRTrig.Q THEN
                    errorFlag := FALSE;
                    state     := IDLE;
                END_IF;
        END_CASE;
    END_IF;

    prev_openBtn  := openBtn;
    prev_closeBtn := closeBtn;
    prev_obstacle := obstacle;
END_FUNCTION_BLOCK

(* CONTRACT_RULES [] *)
